(* IEC 61131-3 sources: daoli-st-library/DL_MathData (part 23) *)

(* ---- FC_DL_SearchMinMaxUdint.st ---- *)
(*
  ==================================================================
  组件名 Component  : FC_DL_SearchMinMaxUdint
  分类   Category   : DL_MathData
  复杂度 Complexity  : 低
  版本   Version    : 1.0.0
  功能   Purpose    : UDINT 域数组单遍扫描求最小值/最大值与双索引同出。前 nCount
                      个元素有效，一次循环同时出 uMin/uMax 与 uMinIdx/uMaxIdx
                      （首命中口径），无效哨兵按开关跳过并计数。
  来源   Source     : t2-1-lgf-math（LGF Math 极值检索族 UDINT 变体）
  溯源   Origin     : 极值检索属公开数学语义，clean-room 自研实现，未复制 LGF
                      或任何厂商私有库源码。
  平台   Platform   : 纯 IEC 61131-3（仅 FOR / 比较 / DINT_TO_UDINT），
                      CODESYS / TwinCAT / InoProShop / Machine Expert 通用
  分工声明 Split     : 与 FC_DL_SearchMinMax（LREAL 属主）及
                      FC_DL_SearchMinMaxDint（DINT 域同批连号件）三角互引——
                      本件为无符号域同构件，判式一律全序（<= / >=），不使用
                      任何减法比较（无符号域差值会回绕成大正数）。
  作者   Author     : 道莅代码库 · PLC 编程专家（R60）
  ------------------------------------------------------------------
  边界 Boundary     :
                      一 扫描个数钳位 1..4096，钳位置信息级码；
                      二 无效样本域：UDINT 域无 NaN，本件无效量定义为哨兵
                         DL_SMU_INVALID（= UDINT 最大位型 16#FFFF_FFFF），仅当
                         bIgnoreInvalid 为真时跳过（与 DINT 件哨兵取最小位型的
                         对称口径，头注释留痕）；
                      三 全量无效时 bValid = FALSE 且双索引回 0，不冒充 0 号位极值；
                      四 无符号比较只允许全序判式 <= / >=，禁用 a - b 差值判序；
                      五 无状态纯函数：每次调用局部量一律段 1 显式预置（R254）。
  接口偏离声明       : 派单示意 fMin/fMax（浮点命名），UDINT 输出按 R265 命名-类型
                      一致性落为 uMin/uMax，语义与引脚数一字不减。
  错误码   Codes    :
    16#0001_0604【信息级】计数越界已钳位（<1 早退，>4096 钳位续扫）
    16#0001_0605【信息级】无效哨兵样本已跳过，个数见 nSkipCnt
    16#0001_0606【故障级】全量无效，无有效极值，bValid = FALSE
  验收   Acceptance :
    算法已证（脚本）：未跑 ｜ 编译器已证（三平台）：未跑
    V1 数据 5 / 3 / 9 / 3，个数 4 → uMin=3 于索引 1，uMax=9 于索引 2
    V2 数据 16#FFFF_FFFE / 0 → uMin=0 于索引 1，uMax=16#FFFF_FFFE 于索引 0
    V3 哨兵 16#FFFF_FFFF 夹在有效值间，bIgnoreInvalid 真 → 跳过 1 个，码含 0605
    V4 个数 0 → bValid=FALSE、码 0604、双索引 0
    V5 全为哨兵且 bIgnoreInvalid 真 → bValid=FALSE、码 0606
  修订记录 Revision  :
    2026-11-21  v1.0.0  R60 首版（批 1 · 序号 2）
  ==================================================================
*)
FUNCTION FC_DL_SearchMinMaxUdint : BOOL
VAR_IN_OUT
    auValues : ARRAY[0..4095] OF UDINT; // 待扫描数组 [计数值]，前 nCount 个有效 / the scanned array, the first nCount entries valid
END_VAR
VAR_INPUT
    nCount         : DINT; // 有效样本数 [个]，钳位 1..4096 / the valid sample count, clamped to one through four thousand ninety six
    bIgnoreInvalid : BOOL; // 是否跳过无效哨兵值 [-] / whether the invalid sentinel entries are skipped
END_VAR
VAR_OUTPUT
    uMin     : UDINT; // 最小值 [计数值]，无有效样本时为 0 / the minimum value, zero when no valid sample
    uMax     : UDINT; // 最大值 [计数值]，无有效样本时为 0 / the maximum value, zero when no valid sample
    uMinIdx  : UDINT; // 最小值所在下标 [下标]，无有效样本时为 0 / the minimum index, zero when no valid sample
    uMaxIdx  : UDINT; // 最大值所在下标 [下标]，无有效样本时为 0 / the maximum index, zero when no valid sample
    nSkipCnt : UDINT; // 被跳过的无效哨兵个数 [个] / the skipped invalid sentinel count
    bValid   : BOOL;  // 结果是否有效（全量无效时为假）[-] / the result validity flag
    eErr     : UDINT; // 错误码，0 = 正常 / the error code, zero is ok
    bError   : BOOL;  // 错误标志，eErr 非 0 时为真 / the error flag, true when eErr is nonzero
END_VAR
VAR
    nI     : DINT;  // 扫描索引 [下标] / the scan index
    nUse   : DINT;  // 钳位后的扫描个数 [个] / the clamped scan count
    nSeen  : DINT;  // 已见有效样本数 [个] / the seen valid sample count
    uV     : UDINT; // 当前样本工作副本 [计数值] / the current sample working copy
    bHave  : BOOL;  // 已取得首个有效样本 [-] / the first valid sample taken flag
    bClamp : BOOL;  // 钳位发生标记 [-] / the clamp happened flag
END_VAR
VAR CONSTANT
    DL_SMU_DMAX    : DINT := 4096;          // 扫描个数上界 [个]，与数组容量一致 / the scan count bound aligned with the array capacity
    DL_SMU_INVALID : UDINT := 16#FFFF_FFFF; // 无效哨兵，等于 UDINT 最大位型（与 DINT 件取最小位型对称）/ the invalid sentinel equal to the UDINT maximum bit pattern
END_VAR

// 段 1｜返回值与错误状态预置安全值（四段式第一段，R45）+ 局部量显式预置（R254）/ segment 1, the preset of the return, the codes and the local guards
FC_DL_SearchMinMaxUdint := FALSE; // 返回值预置假 / preset the return false
uMin := 0; // 最小值预置零 / preset the minimum zero
uMax := 0; // 最大值预置零 / preset the maximum zero
uMinIdx := 0; // 最小索引预置零 / preset the minimum index zero
uMaxIdx := 0; // 最大索引预置零 / preset the maximum index zero
nSkipCnt := 0; // 跳过计数预置零 / preset the skipped count zero
bValid := FALSE; // 有效标志预置假（无有效样本前不宣称有效）/ preset the validity false
eErr := 16#0000_0000; // 错误码预置正常 / preset the code to ok
bError := FALSE; // 错误标志预置假 / preset the error flag false
nUse := 0; // 扫描个数预置零 / preset the scan count zero
nSeen := 0; // 有效样本数预置零 / preset the seen count zero
uV := 0; // 样本工作副本预置零 / preset the sample copy zero
bHave := FALSE; // 首样本标志预置假 / preset the first sample flag false
bClamp := FALSE; // 钳位标记预置假 / preset the clamp flag false

// 段 2｜扫描个数域闸（下界早退 + 上界钳位，边界一）/ segment 2, the scan count domain gate
IF nCount < 1 THEN // 低于下界，无样本可扫 / below the floor, nothing to scan
    eErr := 16#0001_0604; // 信息级：计数越界已钳位 / informational, the count clamped
    bError := TRUE; // 置错误标志（信息级随事件置位惯例）/ raise the error flag
    RETURN; // 早退：bValid 保持 FALSE，双索引保持 0 / early return with the validity false
END_IF
nUse := nCount; // 域内接管 / take the count inside the domain
IF nUse > DL_SMU_DMAX THEN // 高于上界 / above the bound
    nUse := DL_SMU_DMAX; // 钳到数组容量 / clamp to the array capacity
    bClamp := TRUE; // 置钳位标记 / raise the clamp flag
END_IF
IF bClamp THEN // 钳位发生时置信息级 / raise the informational code on a clamp
    eErr := 16#0001_0604; // 信息级：计数越界已钳位 / informational, the count clamped
    bError := TRUE; // 置错误标志 / raise the error flag
END_IF

// 段 3｜单遍扫描：首命中取极小与极大，索引与值同源写出（边界四）/ segment 3, the single pass scan with the first hit rule
FOR nI := 0 TO nUse - 1 DO // 有界循环（nUse 已钳 ≤4096）/ the bounded loop
    uV := auValues[nI]; // 取样本（索引已证在数组界内）/ take the sample, the index proven inside the bounds
    IF bIgnoreInvalid AND (uV >= DL_SMU_INVALID) THEN // 无效哨兵且开关为真（全序判式，不用等号）/ an invalid sentinel with the switch true, a total order test
        nSkipCnt := nSkipCnt + 1; // 跳过计数推进 / advance the skipped count
    ELSE // 有效样本参与极值 / a valid sample participates
        nSeen := nSeen + 1; // 有效样本数推进 / advance the seen count
        IF NOT bHave THEN // 首个有效样本：双向装填 / the first valid sample seeds both sides
            uMin := uV; // 最小值装填 / seed the minimum
            uMax := uV; // 最大值装填 / seed the maximum
            uMinIdx := DINT_TO_UDINT(nI); // 最小索引装填 / seed the minimum index
            uMaxIdx := DINT_TO_UDINT(nI); // 最大索引装填 / seed the maximum index
            bHave := TRUE; // 置首样本标志 / raise the first sample flag
        ELSE // 后续样本比较（首命中用严格判式，不覆盖等值）/ the later samples, strict tests keep the first hit
            IF uV < uMin THEN // 新极小 / a new minimum
                uMin := uV; // 更新最小值 / update the minimum
                uMinIdx := DINT_TO_UDINT(nI); // 更新最小索引（与值同源）/ update the minimum index from the same source
            ELSIF uV > uMax THEN // 新极大（uV ≥ uMin 前提下判极大即可，全序自证）/ a new maximum, proven by the total order
                uMax := uV; // 更新最大值 / update the maximum
                uMaxIdx := DINT_TO_UDINT(nI); // 更新最大索引（与值同源）/ update the maximum index from the same source
            END_IF
        END_IF
    END_IF
END_FOR

// 段 4｜结果复检兜底：全量无效判故障，信息级与故障级不共码（R258 三件套）/ segment 4, the result recheck
IF (nSeen > 0) AND (nSkipCnt > 0) AND (eErr = 16#0000_0000) THEN // 部分跳过且无先发事件 / a partial skip with no earlier event
    eErr := 16#0001_0605; // 信息级：无效哨兵样本已跳过 / informational, the invalid sentinels skipped
    bError := TRUE; // 置错误标志 / raise the error flag
END_IF
IF nSeen < 1 THEN // 无有效样本 / no valid sample
    eErr := 16#0001_0606; // 故障级：全量无效，无有效极值 / fault grade, no valid extremum
    bError := TRUE; // 置错误标志（R45 配对）/ raise the error flag, paired with the fault code
    bValid := FALSE; // 结果不可用 / the result void
    uMin := 0; // 双极值回安全值 / both extrema back to the safe zero
    uMax := 0; // 双极值回安全值 / both extrema back to the safe zero
    uMinIdx := 0; // 索引回 0（不冒充 0 号位极值，边界三）/ the index back to zero, not posing as the entry zero
    uMaxIdx := 0; // 索引回 0（不冒充 0 号位极值，边界三）/ the index back to zero, not posing as the entry zero
ELSE // 有有效样本 / with valid samples
    bValid := TRUE; // 结果有效 / the result is valid
    FC_DL_SearchMinMaxUdint := TRUE; // 返回成功 / return success
END_IF
END_FUNCTION

(* ---- FC_DL_SelEx.st ---- *)
(*
    FC_DL_SelEx —— 双通道选择泛型防御包装（REAL 域）
    ------------------------------------------------------------------
    分类      : DL_MathData / Sel
    前缀      : FC_DL_
    版本      : 1.0.0
    溯源      : IEC 61131-3 标准语义的道莅防御性实现
                （内部委托平台内建函数，外围统一错误码/钳位/双语文档；
                  未复制任何闭源厂商源码，参考实现仅限 MIT/Apache 许可）
    平台      : 纯 IEC 61131-3，CODESYS / TwinCAT / InoProShop 通用
    作者      : 道莅代码库 · PLC编程专家（R16）
    ------------------------------------------------------------------
    功能说明  : 双通道选择：bG=FALSE 选 fI0、bG=TRUE 选 fI1，选择运算用比较与
                IF/ELSE 实现（IEC SEL 语义），不重实现任何数学内核；
                选中通道非有限（NaN 或 ±INF）判为故障级 16#0001_02AC，返回 0.0 且 bValid=FALSE；
                未选中通道（备用通道）非有限仅置信息级 16#0001_01D4 记录，
                不影响本拍输出（输出仍为选中通道的有效值，bError=FALSE、bValid=TRUE）；
                选中与未选中同时异常时，故障级优先（返回 0.0）；
                ±INF 采用平台安全幅值比较判定（阈值高于 REAL 最大有限值 3.402823E38），NaN 用自不等判定；
                钳位方向：无钳位（故障拦截 / 信息记录，输出为通道原值或 0.0）。
    错误码    : 16#0001_02AC 选中通道非有限（NaN 或 ±INF）——故障级，返回 0.0
                16#0001_01D4 未选中通道（备用通道）非有限，仅记录——信息级，不影响本拍输出
                16#0001_01D5 预留禁用（信息级，不得挪用）
                16#0001_02AD 预留禁用（故障级，不得挪用）
                16#0001_02AE 预留禁用（故障级，不得挪用）
    状态机    : R6 标注 N/A —— 本组件为纯函数无顺序状态机，无 CASE 可写，非法状态不可能出现，故以本节说明替代 ELSE 兜底
    修订记录  : 2026-11-16 v1.0.0 首次入库（R16）
*)
FUNCTION FC_DL_SelEx : REAL
VAR_INPUT
    bG  : BOOL; // 选择输入，FALSE 选 fI0、TRUE 选 fI1 / select input, FALSE picks fI0, TRUE picks fI1
    fI0 : REAL; // 通道 0 输入 [无量纲] / channel 0 input
    fI1 : REAL; // 通道 1 输入 [无量纲] / channel 1 input
END_VAR
VAR_OUTPUT
    eErr   : UDINT; // 错误码，0=正常 / error id, 0=ok
    bError : BOOL;  // 是否出错，eErr 非 0 时为 TRUE / error flag, TRUE when eErr is nonzero
    bValid : BOOL;  // 输出是否有效可用 / output valid flag
END_VAR
VAR CONSTANT
    DL_REAL_INF_GUARD : LREAL := 4.0E38; // REAL 域 ±INF 判定阈值，高于 REAL 最大有限值 3.402823E38 [无量纲] / REAL +/-INF guard above max finite REAL 3.402823E38
END_VAR
VAR
    fSel      : REAL; // 选中通道值 [无量纲] / selected channel value
    bSelBad   : BOOL; // 选中通道非有限判定结果 / non-finite detection result of selected channel
    bIdleBad  : BOOL; // 未选中通道非有限判定结果 / non-finite detection result of unselected channel
END_VAR

// 段 1｜返回值与错误状态预置 / segment 1, preset return value and error status
FC_DL_SelEx := 0.0; // 故障缺省返回 0 [无量纲] / fault default returns 0
eErr   := 0;     // 预置无错误 / preset no error
bError := FALSE; // 预置无故障 / preset no fault
bValid := FALSE; // 预置无效，通过防御闸后置位 / preset invalid, set TRUE after guard passes

// 段 2｜通道选择与选中/未选中通道有限性判定 / segment 2, channel selection and finiteness check of both channels
IF bG THEN
    fSel := fI1; // TRUE 选通道 1 / TRUE picks channel 1
    bIdleBad := (fI0 <> fI0) OR (fI0 > DL_REAL_INF_GUARD) OR (fI0 < -DL_REAL_INF_GUARD); // 未选中通道 fI0 非有限判定 [无量纲] / unselected fI0 non-finite check
ELSE
    fSel := fI0; // FALSE 选通道 0 / FALSE picks channel 0
    bIdleBad := (fI1 <> fI1) OR (fI1 > DL_REAL_INF_GUARD) OR (fI1 < -DL_REAL_INF_GUARD); // 未选中通道 fI1 非有限判定 [无量纲] / unselected fI1 non-finite check
END_IF
bSelBad := (fSel <> fSel) OR (fSel > DL_REAL_INF_GUARD) OR (fSel < -DL_REAL_INF_GUARD); // 选中通道非有限判定（NaN 自不等 + 安全幅值判 ±INF） / selected channel non-finite check (NaN by self-inequality, +/-INF by safe magnitude)

// 段 3｜防御闸与输出（末段，故障级优先） / segment 3, guard and output (final, fault level first)
IF bSelBad THEN
    FC_DL_SelEx := 0.0;       // 故障级返回 0 [无量纲] / fault level returns 0
    eErr   := 16#0001_02AC;   // 选中通道非有限故障码 / selected channel non-finite fault id
    bError := TRUE;           // 置故障标志 / set fault flag
    bValid := FALSE;          // 输出无效 / output invalid
    RETURN;                   // 立即返回 / immediate return
ELSIF bIdleBad THEN
    FC_DL_SelEx := fSel;      // 输出选中通道原值，备用通道异常不影响本拍输出 / output selected value, idle channel anomaly does not affect this cycle
    eErr := 16#0001_01D4;     // 信息级：备用通道异常仅记录 / info level: idle channel anomaly recorded only
ELSE
    FC_DL_SelEx := fSel;      // 双通道均有限，正常输出选中值 / both channels finite, normal selected output
    eErr := 0; // 无错误 / no error
END_IF
bError := FALSE; // 信息级记录不置故障，故障分支已提前返回 / info-level record never raises fault, fault branch has returned
bValid := TRUE;  // 选中通道输出有效可用 / selected channel output is valid
END_FUNCTION

(* ---- FC_DL_SignedToUdintSat.st ---- *)
(*
  ==================================================================
  组件名 Component  : FC_DL_SignedToUdintSat
  分类   Category   : DL_MathData
  前缀   Naming     : FC_DL_ ｜ b/n/u/f/t/e/st 类型前缀制（R265）
  码位   Code ID    : 16#0001_0651（信息级）
  版本   Version    : 1.0.0
  复杂度 Complexity  : 低
  功能   Purpose    : DINT → UDINT 确定性转换：负值钳 0 并发信息级提示（多数平台此类
                      隐式转换行为不一，负值可能回绕成巨大正数，是 Modbus 寄存器打包的
                      经典故障源）。
  开源溯源 Origin    : IEC 61131-3 标准语义的道莅防御性实现（clean-room，无第三方代码行）
  许可证 License    : MIT
  参考   Reference  : IEC 61131-3:2013 §6.6.5 类型转换函数与 §6.5 有符号/无符号整数域定义
  平台   Platform   : 纯 IEC 61131-3（DINT_TO_UDINT / 比较），三平台通用
  依赖   Depends    : 仅 Standard.library（DINT_TO_UDINT 属标准转换函数）
  分工声明 Split     : FC_DL_UdintToDintChk 为反方向（UDINT → DINT，超上界钳 MAX 并置
                      故障级码），本件为 DINT → UDINT（负值钳零并置信息级码），两件成对，
                      边界互引（R216）。16 位入口（INT → UINT 同语义）按「禁新增同义邻件」
                      纪律并入本件重载，不另立文件。
  归属 Ownership     : 本件无 TYPE 声明，全部引脚为 IEC 标准原生类型。
  ------------------------------------------------------------------
  边界 Boundary     :
                      一 负值钳零是确定性合法行为而非故障：置信息级码、bValid 保持 TRUE、
                         bError 保持 FALSE（若按故障处理，Modbus 打包遇到合法的负温度
                         就会停机，分级明显错位）；
                      二 正域精确无溢出，域包含证明：DINT 非负域 [0, 2^31 − 1] 是全序
                         子集于 UDINT 全域 [0, 2^32 − 1]，即 [0, 2147483647] ⊂ [0, 4294967295]，
                         故 diIn ≥ 0 时 DINT_TO_UDINT 恒为精确映射，无须溢出分支；
                      三 反方向（UDINT → DINT）的越上界场景在本件域内不可能出现：
                         入参已是 UDINT 域内的值经 DINT 往返，属反方向件职责，本件不设分支；
                      四 纯函数：无记忆量、无定时器、无边沿实例，每调用重算。
  错误码 Codes      :
    16#0001_0651【信息级】负值已钳零（不锁存、不置 bError、bValid 保持 TRUE）
  验收 Acceptance   :
    算法已证（脚本）：未跑 ｜ 编译器已证（三平台）：未跑
    V1 0 → 0、bNegClamped = FALSE、无码
    V2 -1 → 0 + bNegClamped + 码 0651（bError = FALSE）
    V3 MIN（-2147483648）→ 0 + bNegClamped + 码 0651
    V4 MAX（2147483647）→ 2147483647 精确、无码
    V5 反方向向量（2^32−1 入 DINT）域上不可能，注释已给域包含关系，无须代码分支
  修订记录 Revision  :
    2026-11-21  v1.0.0  R62 首版（批 2 · 序号 6）
  ==================================================================
*)
FUNCTION FC_DL_SignedToUdintSat : BOOL
VAR_INPUT
    diIn : DINT; // 有符号输入 [−]，完整 DINT 域 / the signed input over the full DINT domain
END_VAR
VAR_OUTPUT
    udiOut      : UDINT; // 无符号结果 [−] / the unsigned result
    bNegClamped : BOOL;  // 负值已钳零 [-] / a negative value was clamped to zero
    bValid      : BOOL;  // 结果可用（本件恒 TRUE，保留引脚供族内统一）[-] / the result is usable, always true here
    eErr        : UDINT; // 错误码，0 = 正常 / the error code, zero is ok
    bError      : BOOL;  // 故障标志（本件只有信息级码，恒 FALSE）/ the fault flag, always false here since only an informational code exists
END_VAR
VAR CONSTANT
    DL_S2U_ZERO : DINT := 0;                  // 有符号零常量 [−] / the signed zero constant
    DL_S2U_UMIN : UDINT := 0;                 // 无符号零常量 [−] / the unsigned zero constant
    DL_S2U_DMAX : DINT := 2147483647;         // DINT 可表达上界 [−]，即 2^31−1 / the expressible DINT ceiling, two to the thirty first minus one
    DL_S2U_UMAX : UDINT := 4294967295;        // UDINT 可表达上界 [−]，即 2^32−1 / the expressible UDINT ceiling, two to the thirty second minus one
END_VAR

// 段 1｜返回值与全部出口预置安全值（R45 四段式第一段）/ segment 1, preset every outlet to its safe value
FC_DL_SignedToUdintSat := FALSE; // 返回值预置假 / preset the return false
udiOut := DL_S2U_UMIN; // 结果预置零 [−] / preset the result zero
bNegClamped := FALSE; // 负值钳零标志预置假 / preset the negative clamp flag false
bValid := FALSE; // 可用标志预置假，过闸后置位 / preset the validity false, raised after the gates
eErr := 16#0000_0000; // 错误码预置正常 / preset the code to ok
bError := FALSE; // 故障标志预置假（本件无故障级码）/ preset the fault flag false, no fault level code exists here

// 段 2｜负值钳零（边界一：确定性行为，非故障）/ segment 2, the negative clamp is a deterministic behaviour, not a fault
IF diIn < DL_S2U_ZERO THEN // 负值域 / the negative domain
    udiOut := DL_S2U_UMIN; // 钳零 [−] / clamp to zero
    bNegClamped := TRUE; // 置钳零标志 / raise the negative clamp flag
    eErr := 16#0001_0651; // 信息级：负值已钳零 / informational, a negative value was clamped to zero
    bError := FALSE; // 明确不置故障标志（信息级，R285 分级纪律）/ keep the fault flag false, this is informational
ELSE // 非负域：精确映射（边界二域包含证明）/ the non negative domain maps exactly
    udiOut := DINT_TO_UDINT(diIn); // 标准显式转换（DINT 非负域 ⊆ UDINT 全域）[−] / the standard explicit conversion, the signed non negative domain is a subset of the unsigned domain
END_IF

// 段 3｜统一出口（信息级钳零仍可用）/ segment 3, the unified outlet where a clamped zero stays usable
bValid := TRUE; // 负值钳零与正域精确均可用 / both the clamped zero and the exact positive domain are usable
FC_DL_SignedToUdintSat := TRUE; // 返回成功 / return success
END_FUNCTION

(* ---- FC_DL_SignumCalc.st ---- *)
(*
    FC_DL_SignumCalc —— 三态符号函数（浮点容差判零 + 非有限拦截）
    ------------------------------------------------------------------
    分类      : DL_MathData / Math-Sign
    前缀      : FC_DL_
    版本      : 1.0.0
    来源标签  : iec-std-wrapper（T0）
    溯源      : IEC 61131-3 标准语义的道莅防御性实现
                （纯比较逻辑，无内建数学内核依赖；未复制任何闭源厂商源码）
    平台      : 纯 IEC 61131-3，CODESYS / TwinCAT / InoProShop 通用
    分工声明  : 与存量 FC_DL_RealEqTolEx（判等）分工——EqTolEx 只回答是否相等，
                本件返回三态符号（负/零/正）；与 Hysteresis 分工——迟滞件带
                状态记忆，本件为无状态纯函数。
    作者      : 道莅代码库 · PLC 编程专家（R57）
    ------------------------------------------------------------------
    功能说明  : 返回输入的三态符号：|x| < fEps 判零返回 0（禁 = 判等）；
                x <= -fEps 返回 -1；x >= fEps 返回 +1。fEps <= 0 组态错误
                返回 0；非有限（NaN/Inf 双判据）返回 0 并出错误码。
    错误码    : 0000 正常 / 16#0003_0001 入参非有限 / 16#0003_0002 fEps 组态非法
    修订记录  : 2026-11-21 v1.0.0 首次入库（R57 批 3 · 序号 11）
*)
FUNCTION FC_DL_SignumCalc : INT
VAR_INPUT
    lrIn : LREAL;       // 输入实数 [工程单位] / input real value [engineering unit]
    fEps : LREAL := 1E-9; // 判零容差 [工程单位]，域 大于零 / the zero tolerance [engineering unit], above zero
END_VAR
VAR_OUTPUT
    eErr   : UDINT; // 错误码，0 = 正常 / error code, zero is ok
    bError : BOOL;  // 出错标志，eErr 非 0 时为真 / error flag, true when eErr is nonzero
    bValid : BOOL;  // 结果是否可用，拦截/组态错误时为假 / the result usable, false when intercepted
END_VAR

// 段 1｜返回值与错误状态预置安全值（四段式第一段，R45）/ segment 1, preset the return and error states
FC_DL_SignumCalc := 0; // 符号预置零 / preset the sign to zero
eErr   := 16#0000_0000; // 错误码预置正常 / preset the code to ok
bError := FALSE; // 错误标志预置假 / preset the error flag false
bValid := TRUE; // 有效标志预置真 / preset the valid flag true

// 段 2｜非有限拦截（双判据）：命中早退不比较 / segment 2, the non finite interception
IF (lrIn <> lrIn) OR ((lrIn - lrIn) <> (lrIn - lrIn)) THEN // NaN 或无穷 / NaN or infinity
    eErr   := 16#0003_0001; // 信息级：输入非有限返回零 / informational, a non finite input returns zero
    bError := TRUE; // 置错误标志 / raise the error flag
    bValid := FALSE; // 输出不可用 / the output void
    RETURN; // 返回预置安全值 0 / return the preset safe zero
END_IF

// 段 3｜组态闸：fEps <= 0 判组态错误（边界十一）/ segment 3, the config gate, a nonpositive tolerance illegal
IF (fEps <= 0.0) OR (fEps <> fEps) OR ((fEps - fEps) <> (fEps - fEps)) THEN // 容差非法或非有限 / an illegal or non finite tolerance
    eErr   := 16#0003_0002; // 错误级：容差组态非法 / error grade, an illegal tolerance config
    bError := TRUE; // 置错误标志 / raise the error flag
    bValid := FALSE; // 输出不可用 / the output void
    RETURN; // 返回预置安全值 0 / return the preset safe zero
END_IF

// 段 4｜三态符号判定：容差判零，禁 = 判等（边界十一）/ segment 4, the three state verdict with the tolerance
IF lrIn >= fEps THEN // 显著为正 / clearly positive
    FC_DL_SignumCalc := 1; // 返回正号 / return plus one
ELSIF lrIn <= -fEps THEN // 显著为负 / clearly negative
    FC_DL_SignumCalc := -1; // 返回负号 / return minus one
ELSE // 容差带内判零 / inside the tolerance band
    FC_DL_SignumCalc := 0; // 返回零 / return zero
END_IF
END_FUNCTION

(* ---- FC_DL_SimpsonQuad.st ---- *)
(*==============================================================================
 * 组件名称 (Component)  : FC_DL_SimpsonQuad
 * 所属子库 (Sublibrary) : DL_MathData
 * 当前版本 (Version)    : 1.0.0
 * 兼容性   (Platform)   : CODESYS 3.5+ / TwinCAT 3 / 汇川 InoProShop / 施耐德 Machine Expert
 *                         仅依赖 Standard.library（LOWER_BOUND / UPPER_BOUND / MOD），零厂商私有库
 * 功能描述 (Function)   : 复合辛普森 1/3 数值积分原语：对 n+1 个等距节点纵坐标（n 为偶数，
 *                         即节点数 >= 3 且区间数为偶）按公式
 *                           fI = fDx/3 × (aY[0] + 4×Σ奇节点 + 2×Σ偶内点 + aY[n])
 *                         单遍求积，返回积分值。适用功率-时间曲线求能、流量累计复核等
 *                         叶子级数值积分场景。
 * 接口     (Interface)  : 输入 aY 等距节点纵坐标数组（变长数组，按引传）、fDx 节点步长；
 *                         引用输出 bValid 有效标志（REFERENCE TO BOOL，当拍写回）；
 *                         返回值 = 积分值（bValid=FALSE 时返回 0）。
 * 边界     (Boundary)   : ① **属主边界（写死）：本件只做一次静态数组求积，不采样、不缓存、
 *                         不做时间触发**；采样与节点装载由调用方负责。
 *                         ② 奇偶判据用整数 MOD 2，禁浮点判奇偶。
 *                         ③ 拒算条件（任一成立返回 0 且 bValid=FALSE）：区间数 < 2（节点数
 *                         < 3）、区间数为奇数、fDx <= 容差、任一节点纵坐标非有限
 *                         （NaN 用自不等 x<>x 口径、Inf 用 (x-x)<>0 口径，R245）。
 *                         非有限值逐点前置剔除并**整体拒算**：部分积分结果不可信。
 *                         ④ 等距性由调用方保证（IN 语义声明）：本件不做步长一致性校验，
 *                         fDx 取相邻节点间距的名义值。
 *                         ⑤ 变长数组仅入 VAR_IN_OUT（IEC 61131-3 第 3 版对 ARRAY[*] 的
 *                         传参域限定），LOWER_BOUND/UPPER_BOUND 取实际上下界，不假设 0 起始。
 *                         ⑥ 零全局耦合（无 GVL / 无 VAR_EXTERNAL / 无物理地址）。
 * 分工声明 (Scope)      : 与 `FC_DL_PolyEvalHorner` 分工：多项式求值 ≠ 数值求积；与
 *                         `FC_DL_MultiPointLinear` 分工：分段线性插值 ≠ 积分。全库数值
 *                         积分原语由本件开族。
 * 来源标签 (Source Tag) : T2-1 LGF · Math 数学子族（公开数学定义 clean-room，复合辛普森
 *                         1/3 法则为教科书公开公式，零代码行复制）
 * 码表     (Codes)      : 本件不占用任何全局数字码位。出口为 LREAL 积分值 + BOOL 有效标志；
 *                         数字码位待主控收口阶段统一派号。
 * 红线自检 (Redline)    : R1 ✓ 零 GVL/VAR_EXTERNAL ｜ R2 ✓ 零 %I/%Q/%M ｜ R3 ✓ 纯 IEC 61131-3
 *                         R4 ✓ 步长容差闸 + 非有限前置剔除 + 奇偶整数判据 ｜ R5 ✓ 声明逐行同行双语注释
 *                         R6 N/A（纯函数无状态机） ｜ R7 N/A（无实例调用）
 * 修订历史 (Revision)   : 2026-11-20  v1.0.0  R48 首版（批次 1 · 序号 2）
 *                         验收向量：3 节点 y=[0,1,0]、dx=1 → 4/3；4 节点（奇区间数）拒算；
 *                         含 NaN 节点整体拒算；dx=0 拒算。
 *==============================================================================*)

FUNCTION FC_DL_SimpsonQuad : LREAL
VAR_IN_OUT
    aY : ARRAY[*] OF LREAL;    // 等距节点纵坐标数组（长度 n+1，n 偶），单位随被积量 [被积量纲] / Ordinates at equidistant nodes
END_VAR
VAR_INPUT
    fDx    : LREAL;                 // 节点步长，域 > 容差；等距性由调用方保证（IN 语义） [横轴单位] / Node spacing, > epsilon, uniformity by caller
    bValid : REFERENCE TO BOOL;     // 有效标志（引用传参；FALSE=拒算） [-] / Validity flag, by-reference, FALSE when rejected
END_VAR
VAR
    nLo  : DINT;                    // 数组实际下界索引 / Actual lower array index
    nHi  : DINT;                    // 数组实际上界索引 / Actual upper array index
    nInt : DINT;                    // 区间数 = 节点数 - 1，须为正偶数 / Interval count, positive even
    i    : DINT;                    // 求和循环索引 / Summation loop index
    fSum : LREAL;                   // 括号内加权和中间量 / Weighted sum accumulator
END_VAR
VAR CONSTANT
    DL_SQ_EPS : LREAL := 1.0E-12;   // 步长判零容差 [横轴单位] / Spacing zero epsilon
    DL_SQ_W4  : LREAL := 4.0;       // 辛普森奇节点权重 [-] / Simpson odd-node weight
    DL_SQ_W2  : LREAL := 2.0;       // 辛普森偶内点权重 [-] / Simpson even-interior weight
    DL_SQ_W3  : LREAL := 3.0;       // 1/3 法则除数 [-] / Divisor of the one-third rule
END_VAR

bValid := FALSE;                                       // 缺省拒算 / Default: invalid
FC_DL_SimpsonQuad := 0.0;                              // 拒算返回 0 / Rejected returns zero
nLo  := LOWER_BOUND(aY, 1);                            // 取实际下界，不假设 0 起始 / Actual lower bound, no zero assumption
nHi  := UPPER_BOUND(aY, 1);                            // 取实际上界 / Actual upper bound
nInt := nHi - nLo;                                     // 区间数 / Interval count
IF (nInt < 2) OR ((nInt MOD 2) <> 0) OR (fDx <= DL_SQ_EPS) THEN
    RETURN;                                            // 区间数不足 / 奇区间数 / 步长非正：拒算（整数奇偶判据）/ Too few or odd intervals or bad spacing: reject
END_IF
FOR i := nLo TO nHi DO
    IF (aY[i] <> aY[i]) OR ((aY[i] - aY[i]) <> 0.0) THEN
        RETURN;                                        // 任一节点非有限（NaN 自不等 / Inf 差非零）：整体拒算（R245）/ Any non-finite node: reject wholly
    END_IF
END_FOR

fSum := aY[nLo] + aY[nHi];                             // 两端节点权重 1 / End nodes carry weight one
FOR i := (nLo + 1) TO (nHi - 1) DO
    IF ((i - nLo) MOD 2) <> 0 THEN
        fSum := fSum + DL_SQ_W4 * aY[i];               // 奇节点权重 4 / Odd nodes weight four
    ELSE
        fSum := fSum + DL_SQ_W2 * aY[i];               // 偶内点权重 2 / Even interior nodes weight two
    END_IF
END_FOR

FC_DL_SimpsonQuad := fSum * fDx / DL_SQ_W3;            // 除数为常量 3，无除零 / Constant divisor three, no zero division
bValid := TRUE;                                        // 求积有效 / Result valid

END_FUNCTION

(* ---- FC_DL_SincSafe.st ---- *)
(*==============================================================================
 * 名称 : FC_DL_SincSafe —— 安全 sinc(x)=sin(x)/x（0 点泰勒展开防除零）
 * 分类 / 前缀 / 版本 : DL_MathData / FC_DL_ / 1.0.0
 * 溯源 : 开源语义参考（OSCAT/AixOCAT 族，MIT）或 clean-room IEC 实现，未复制源码
 * 平台 : 纯 IEC 61131-3
 * 功能说明 : 计算 sinc(x)=sin(x)/x。|x|<1.0E-8 时用四阶泰勒近似
 *            1 - x^2/6 + x^4/120（该区间误差 < 1.0E-16 量级），避免 0 点
 *            除零；其余区间直接 sin(x)/x（|x|>=1.0E-8 保证分母非零）。
 *            边界处理：输入非有限（NaN/±Inf）置 eErr 返回 0.0；x=0 精确落
 *            入泰勒支路返回 1.0（sinc 极限值），属正确结果非故障。
 * 错误码 : 16#0001_1B0F = 输入非有限（NaN/±Inf）
 *          eErr=0 且 bValid=TRUE 表示返回值可用
 * 状态机 : R6 标注 N/A（纯函数无顺序状态，以本节替代 ELSE 兜底）
 * 红线 : R1/R2/R3 ✓ 零全局/零IO/纯IEC ｜ R4 ✓ 非有限拦截/除零防护 ｜ R10 ✓ 标准转换 ｜ R11 ✓ 分号收尾 ｜ R15 ✓ 无保留字撞名
 * 修订记录 : 2026-11-23 v1.0.0 首次入库（R76）
 *============================================================================*)
FUNCTION FC_DL_SincSafe : LREAL
VAR_INPUT
    fX : LREAL;    // 输入自变量 [rad] / input argument in radians
END_VAR
VAR_OUTPUT
    eErr   : UDINT;    // 故障码，0=正常，1B0F=输入非有限 / error code
    bError : BOOL;     // TRUE=本件发生故障 / TRUE when fault occurred
    bValid : BOOL;     // TRUE=返回值可用 / TRUE when return value is usable
END_VAR
VAR
    _x2 : LREAL;       // x 的平方（泰勒中间量）/ squared input for Taylor series
    _x4 : LREAL;       // x 的四次方（泰勒中间量）/ fourth power for Taylor series
END_VAR

FC_DL_SincSafe := 0.0;                       // 返回值预设 0.0 / preset return to zero
eErr   := 16#0000_0000;                      // 故障码清零 / clear error code
bError := FALSE;                             // 故障标志清零 / clear error flag
bValid := TRUE;                              // 预设输出可用 / preset valid flag

IF (fX <> fX) OR ((fX - fX) <> (fX - fX)) THEN    // NaN 或 ±Inf / NaN or infinite
    eErr   := 16#0001_1B0F;                  // 置非有限故障码 / set non-finite code
    bError := TRUE;                          // 置故障标志 / set error flag
    bValid := FALSE;                         // 返回值不可用 / return not usable
    RETURN;                                  // 返回 0.0 / return zero
END_IF

IF ABS(fX) < 1.0E-8 THEN                     // 0 点邻域走泰勒支路 / Taylor branch near zero
    _x2 := fX * fX;                          // 平方中间量 / square
    _x4 := _x2 * _x2;                        // 四次方中间量 / fourth power
    FC_DL_SincSafe := 1.0 - _x2 / 6.0 + _x4 / 120.0;    // 四阶泰勒近似（0 点返回 1.0）/ 4th-order Taylor
ELSE                                         // 非零区间直接作商（分母 |x|>=1E-8 非零）/ direct quotient
    FC_DL_SincSafe := SIN(fX) / fX;          // sin(x)/x，分母已保证非零 / denominator guaranteed nonzero
END_IF

END_FUNCTION

(* ---- FC_DL_SinDeg.st ---- *)
(*==============================================================================
 * 名称 : FC_DL_SinDeg —— 角度制正弦（度入参，弧度内部换算）
 * 分类 / 前缀 / 版本 : DL_MathData / FC_DL_ / 1.0.0
 * 溯源 : 开源语义参考（OSCAT/AixOCAT 族，MIT）或 clean-room IEC 实现，未复制源码
 * 平台 : 纯 IEC 61131-3
 * 功能说明 : 返回 sin(fDeg)：内部换算弧度 fDeg * PI / 180 后调用标准 SIN，
 *            PI 取 LREAL 字面量 3.14159265358979323846（双精度最近舍入）。
 *            边界处理：输入非有限（NaN：f<>f；±Inf：(f-f)<>(f-f)）置 eErr
 *            返回 0.0；|fDeg|>1.0E12 时大角换算精度塌陷，同置 eErr 返回 0.0。
 * 错误码 : 16#0001_1B09 = 输入非有限（NaN/±Inf）或角度量超安全量程 ±1.0E12
 *          eErr=0 且 bValid=TRUE 表示返回值可用
 * 状态机 : R6 标注 N/A（纯函数无顺序状态，以本节替代 ELSE 兜底）
 * 红线 : R1/R2/R3 ✓ 零全局/零IO/纯IEC ｜ R4 ✓ 非有限拦截/量程防护 ｜ R10 ✓ 标准转换 ｜ R11 ✓ 分号收尾 ｜ R15 ✓ 无保留字撞名
 * 修订记录 : 2026-11-23 v1.0.0 首次入库（R76）
 *============================================================================*)
FUNCTION FC_DL_SinDeg : LREAL
VAR_INPUT
    fDeg : LREAL;    // 输入角 [度] / input angle in degrees
END_VAR
VAR_OUTPUT
    eErr   : UDINT;    // 故障码，0=正常，1B09=输入非有限或超量程 / error code
    bError : BOOL;     // TRUE=本件发生故障 / TRUE when fault occurred
    bValid : BOOL;     // TRUE=返回值可用 / TRUE when return value is usable
END_VAR

FC_DL_SinDeg := 0.0;                         // 返回值预设 0.0 / preset return to zero
eErr   := 16#0000_0000;                      // 故障码清零 / clear error code
bError := FALSE;                             // 故障标志清零 / clear error flag
bValid := TRUE;                              // 预设输出可用 / preset valid flag

IF (fDeg <> fDeg) OR ((fDeg - fDeg) <> (fDeg - fDeg))    // NaN 或 ±Inf / NaN or infinite
   OR (ABS(fDeg) > 1.0E12) THEN              // 超安全量程（精度塌陷防护）/ beyond safe range
    eErr   := 16#0001_1B09;                  // 置故障码 / set error code
    bError := TRUE;                          // 置故障标志 / set error flag
    bValid := FALSE;                         // 返回值不可用 / return not usable
    RETURN;                                  // 返回 0.0 / return zero
END_IF

FC_DL_SinDeg := SIN(fDeg * 3.14159265358979323846 / 180.0);    // 度转弧度后取正弦 / degrees to radians, then sine

END_FUNCTION

(* ---- FC_DL_SinEx.st ---- *)
(*
    FC_DL_SinEx —— 正弦防御包装（2π 周期归约保精度 + 非有限拦截 + 超大角度降级）
    ------------------------------------------------------------------
    分类      : DL_MathData / Math-Trig
    前缀      : FC_DL_
    版本      : 1.0.0
    溯源      : IEC 61131-3 标准语义的道莅防御性实现
                （内部委托平台内建函数，外围统一错误码/钳位/双语文档；
                  未复制任何闭源厂商源码，参考实现仅限 MIT/Apache 许可）
    平台      : 纯 IEC 61131-3，CODESYS / TwinCAT / InoProShop 通用
    作者      : 道莅代码库 · PLC编程专家（R15）
    ------------------------------------------------------------------
    功能说明  : 求输入弧度的正弦值。入口先做非有限拦截（NaN/Inf 返回 0.0
                并置 16#0001_0163）；随后按 2π 做周期归约，商取 FLOOR 语义避免负向
                误差，商绝对值 < 2.0E9 保证 DINT 转换不溢出；超大角度
                （绝对值 > 1.0E12 或商超 DINT 安全域）降级处理：置 16#0001_0163、
                bValid=FALSE 但仍继续计算；域内委托内建 SIN，结果再做
                NaN 复检兜底，全程不输出 NaN/Inf。
    错误码    : 0000 正常 / 16#0001_0163 入参越界（非有限输入或超大角度降级，已归零/降级可用）
    修订记录  : 2026-11-16 v1.0.0 首次入库（R15）
*)
FUNCTION FC_DL_SinEx : LREAL
VAR_INPUT
    lrRad : LREAL; // 输入角度 [rad]，任意有限弧度值 / input angle [rad], any finite radian value
END_VAR
VAR_OUTPUT
    eErr : UDINT; // 错误码，0=正常，1=入参越界（非有限或超大角度） / error id, 0=ok, 1=input out of domain (non-finite or super-large angle)
    bError   : BOOL; // 是否出错，eErr 非 0 时为 TRUE / error flag, TRUE when eErr is nonzero
    bValid   : BOOL; // 输出是否有效可用，超大角度降级时为 FALSE / output valid, FALSE for degraded super-large angle
END_VAR
VAR
    lrQ   : LREAL; // 周期商 [周期数]，输入角除以 2π / cycle quotient [cycles], input divided by two pi
    nCyc  : DINT; // 归约周期数 [周期数]，FLOOR 语义整数 / reduction cycle count [cycles], integer with floor semantics
    lrRed : LREAL; // 归约后弧度 [rad]，域约至 0 到 2π / reduced angle [rad], bounded to 0 to 2 pi
END_VAR
VAR CONSTANT
    DL_SN_MAXREAL : LREAL := 1.7976931348623157E308; // 双精度有限极值 [rad]，超界判无穷 / double precision finite max [rad], beyond treated as infinity
    DL_SN_TWOPI   : LREAL := 6.283185307179586; // 圆周率两倍 [rad]，归约模数 / two pi [rad], reduction modulus
    DL_SN_BIG     : LREAL := 1.0E12; // 超大角度阈值 [rad]，超过判降级 / super-large angle threshold [rad], beyond degraded
    DL_SN_QMAX    : LREAL := 2.0E9; // 周期商安全域 [周期数]，保证 DINT 转换不溢出 / quotient safe bound [cycles], keeps DINT conversion overflow-free
    DL_SN_EPS     : LREAL := 1.0E-9; // 浮点容差 [无量纲] / floating point tolerance [dimensionless]
END_VAR

// 段 1｜返回值与错误状态预置，任何早退路径不留脏码 / segment 1, preset return value and error states
FC_DL_SinEx := 0.0; // 返回值预置安全值 0.0 / preset return to safe value 0.0
eErr    := 16#0000_0000; // 错误码预置正常 / preset error id to ok
bError      := FALSE; // 错误标志预置无错 / preset error flag to FALSE
bValid      := TRUE; // 有效标志预置可用 / preset valid flag to TRUE

// 段 2｜非有限拦截：NaN 用自不等判据，无穷用超极值判据 / segment 2, non-finite interception
IF (lrRad <> lrRad) OR (lrRad > DL_SN_MAXREAL) OR (lrRad < -DL_SN_MAXREAL) THEN
    eErr := 16#0001_0163; // 信息级：输入非有限，已归零 / informational, non-finite input, zeroed
    bError   := TRUE; // 置错误标志 / raise error flag
    bValid   := FALSE; // 输出不可用 / output invalid
    RETURN; // 返回预置安全值 0.0 / return preset safe value 0.0
END_IF

// 段 3｜2π 周期归约（FLOOR 语义）：商超 DINT 安全域则跳过归约原值直通 / segment 3, two-pi reduction with floor semantics, skipped when quotient exceeds the DINT safe bound
lrQ := lrRad / DL_SN_TWOPI; // 周期商 [周期数] / cycle quotient [cycles]
IF ABS(lrQ) < DL_SN_QMAX THEN
    nCyc := TRUNC(lrQ); // 向零截取周期数 / truncate quotient toward zero
    IF (lrQ < 0.0) AND (ABS(lrQ - DINT_TO_LREAL(nCyc)) > DL_SN_EPS) THEN
        nCyc := nCyc - 1; // 负非整数商补一，落实 FLOOR 语义 / decrement for negative non-integer quotient to enforce floor semantics
    END_IF
    lrRed := lrRad - DL_SN_TWOPI * DINT_TO_LREAL(nCyc); // 归约后弧度 [rad] / reduced angle [rad]
ELSE
    lrRed := lrRad; // 商超安全域，放弃归约原值直通 / quotient beyond safe bound, reduction skipped
END_IF

// 段 4｜超大角度精度闸：置 16#0001_0163 降级但继续计算 / segment 4, super-large angle precision gate, degraded with code 1 but computation continues
IF (ABS(lrRad) > DL_SN_BIG) OR (ABS(lrQ) >= DL_SN_QMAX) THEN
    eErr := 16#0001_0163; // 信息级：超大角度，精度不可保证 / informational, super-large angle, precision not guaranteed
    bError   := TRUE; // 置错误标志 / raise error flag
    bValid   := FALSE; // 降级输出，需上层注意 / degraded output, upper layer attention required
END_IF

// 段 5｜委托内建 SIN + 结果 NaN 复检兜底 / segment 5, delegation to built-in SIN with result NaN recheck
FC_DL_SinEx := SIN(lrRed); // 委托内建 SIN 内核，不自实现三角内核 / delegate to built-in SIN kernel
IF FC_DL_SinEx <> FC_DL_SinEx THEN
    FC_DL_SinEx := 0.0; // 兜底安全值 / bottom-line safe value
    IF eErr = 16#0000_0000 THEN
        eErr := 16#0001_0163; // 首事件优先置码 / first-event priority code
        bError   := TRUE; // 置错误标志 / raise error flag
        bValid   := FALSE; // 输出不可用 / output invalid
    END_IF
END_IF
END_FUNCTION

(* ---- FC_DL_SinterShrinkageCalc.st ---- *)
(*
  Component : FC_DL_SinterShrinkageCalc
  Category  : DL_MathData
  Type      : FC
  Complexity: C1
  VERSION   : v1.0.0
  功能      : 烧结线收缩率与模具尺寸补偿：按烧结前后密度比开立方得线收缩率，并由成品尺寸反算所需模具尺寸。
  开源溯源  : 道莅原创 clean-room 自研（无外部代码引用）｜License: MIT
  边界条件  : ① 生坯密度与烧结密度均须 > 1e-9（均为除子），否则返回哨兵 -1；
              ② 烧结密度低于生坯密度时收缩率为负（膨胀），照实输出不钳位，便于诊断工艺异常；
              ③ 反算模具尺寸用 成品尺寸 / 线性比例因子，比例因子为 0 时不计算。
*)
FUNCTION FC_DL_SinterShrinkageCalc : REAL
VAR_INPUT
    fGreenDensGcm3 : REAL;   (* 烧结前生坯密度 [g/cm³] Green density before sintering *)
    fSinterDensGcm3: REAL;   (* 烧结后密度 [g/cm³] Sintered density *)
    fFinalDimMm    : REAL;   (* 成品目标尺寸 [mm] Final part dimension *)
END_VAR
VAR_OUTPUT
    fLinFactor  : REAL;   (* 线性比例因子（成品/模具） [-] Linear scale factor *)
    fShrinkPct  : REAL;   (* 线收缩率 [%] Linear shrinkage percent *)
    fDieDimMm   : REAL;   (* 反算模具尺寸 [mm] Die dimension *)
    xValid      : BOOL;   (* 计算有效性标志 [-] Calculation valid flag *)
END_VAR
VAR CONSTANT
    DL_EPS      : REAL := 1.0E-9;   (* 除零判定容差 [无量纲] Divide-by-zero tolerance *)
    DL_THIRD    : REAL := 0.3333333333333333;  (* 立方根指数 [-] Cube-root exponent *)
    DL_PCT_BASE : REAL := 100.0;    (* 百分比基准 [%] Percent base *)
    DL_ONE      : REAL := 1.0;      (* 单位常数 [-] Unity constant *)
END_VAR
(* 出口预置：三出口统一预置 *)
fLinFactor := 1.0; fShrinkPct := 0.0; fDieDimMm := 0.0; xValid := FALSE;
(* 非有限拦截：自反判 NaN，自身差值判 Inf *)
IF (fGreenDensGcm3 <> fGreenDensGcm3) OR ((fGreenDensGcm3 - fGreenDensGcm3) <> 0.0)
   OR (fSinterDensGcm3 <> fSinterDensGcm3) OR ((fSinterDensGcm3 - fSinterDensGcm3) <> 0.0)
   OR (fFinalDimMm <> fFinalDimMm) OR ((fFinalDimMm - fFinalDimMm) <> 0.0) THEN
    FC_DL_SinterShrinkageCalc := -1.0;  (* 哨兵 -1：输入非有限 / Sentinel -1 non-finite *)
    RETURN;
END_IF
(* 组态域闸：两个密度均为除子，成品尺寸须为正 *)
IF (fGreenDensGcm3 <= DL_EPS) OR (fSinterDensGcm3 <= DL_EPS) OR (fFinalDimMm <= DL_EPS) THEN
    FC_DL_SinterShrinkageCalc := -1.0;  (* 哨兵 -1：组态非法 / Sentinel -1 bad config *)
    RETURN;
END_IF
(* 质量守恒：体积比 = 密度比的反比，线比例因子 = 体比例因子的立方根 *)
fLinFactor := EXPT(fGreenDensGcm3 / fSinterDensGcm3, DL_THIRD);
(* 线收缩率：收缩为正，膨胀为负，照实输出便于工艺诊断 *)
fShrinkPct := (DL_ONE - fLinFactor) * DL_PCT_BASE;
(* 反算模具尺寸：成品 = 模具 × 线比例因子，因子为 0 时不下发 *)
IF fLinFactor > DL_EPS THEN
    fDieDimMm := fFinalDimMm / fLinFactor;
END_IF
xValid := TRUE;                            (* 链路有效 / Chain valid *)
FC_DL_SinterShrinkageCalc := fShrinkPct;   (* 返回线收缩率 [%] / Return linear shrinkage *)
END_FUNCTION

(* ---- FC_DL_SlewRateCalc.st ---- *)
(*
  ==================================================================
  组件名 Component  : FC_DL_SlewRateCalc
  分类   Category   : DL_MathData
  前缀   Naming     : FC_DL_ ｜ b/n/u/f 类型前缀制（R265）
  版本   Version    : 1.0.0
  功能   Purpose    : 采样间变化率：fRate = (fCurVal − fPrevVal) / fDtSec
                      [工程单位/s]。fDtSec ≤ 0 闸（除法前置，含容差判零
                      语义：≤0 即拒）；输入非有限闸；差值/结果非有限复
                      核（有限大数相减可溢出 Inf）。纯无状态函数，采样
                      时刻由调用方维护（前后两次采样值由调用方快照传入），
                      本件不驻留上拍数据。
  来源   Source     : t2-1-lgf-technology（差分变化率为公开数值口径，
                      实现零源码复制）
  互引   Cross-ref  : FB_DL_CycleTimeMeasure（同族周期测量件：其扫描周期
                      口径可作 fDtSec 注入来源）；FC_DL_NormTo01（同族
                      数学原子邻件）
  平台   Platform   : 纯 IEC 61131-3 四则 + ABS，三平台通用
  依赖   Depends    : 无 DL_ 内部依赖；无标准库
  红线   Redline    : R1 零全局/VAR_EXTERNAL/R2 零 %I/%Q/R3 纯 IEC 标准
                      R4 除零闸（dt ≤ 0 前置）+ 非有限三面闸（输入/差值/
                      结果）/R5 全变量双语同行注释/R6 纯函数无状态机
                      （CASE 不适用）/R7 无定时器与沿检测/R8 容差常量化
  错误码 Codes      : 01【失效级】采样间隔非法（fDtSec ≤ 0），返回 0
                      02【失效级】任一输入非有限（NaN 自反判 / Inf 上限
                      兜底判）或差值/结果非有限，返回 0
  码位反证 Note     : 01/02 分立依据（R90）：01 在时基面（调用方采样节拍
                      组态/断拍）、02 在数据面可观测；02 若并入 01，则
                      「时基正常仍失败」的数据病态将不可观测，故必须分立。
  验收   Acceptance : V1 10→12 / dt=0.5s → 4 [u/s] ｜ V2 dt=0 → 码 01
                      ｜ V3 dt=−1 → 码 01 ｜ V4 含 NaN → 码 02 ｜
                      V5 1E308→−1E308 / dt=1 → 码 02（差值 Inf）
  变更   Revision   : 2026-11-22  v1.0.0  R67 首版（编码阶段批 2 序 4）
  ==================================================================
*)
FUNCTION FC_DL_SlewRateCalc : LREAL
VAR_INPUT
    fCurVal  : LREAL;  // 当前采样值 [工程单位] / the current sample value
    fPrevVal : LREAL;  // 前一采样值（调用方快照）[工程单位] / the previous sample value, snapshot by the caller
    fDtSec   : LREAL;  // 采样间隔 [s]，须 > 0 / the sample interval in seconds, must be positive
END_VAR
VAR_OUTPUT
    bValid : BOOL;     // 变化率可用标志 [-] / the slew rate usable flag
    nErrId : UDINT;    // 错误码，0=正常，01/02 见头注 [码] / the error code [code]
END_VAR
VAR
    fDelta : LREAL;    // 差值工作寄存器 [工程单位] / the delta working register
END_VAR
VAR CONSTANT
    SRC_FIN_MAX  : LREAL := 1.7976931348623157E308; // LREAL 有限上限 / the finite LREAL limit
    SRC_ERR_NONE : UDINT := 16#0000_0000;           // 无错误 [码] / no error [code]
    SRC_ERR_DT   : UDINT := 16#0000_0001;           // 码 01：采样间隔非法 / code 01, illegal interval
    SRC_ERR_NAN  : UDINT := 16#0000_0002;           // 码 02：非有限 / code 02, non finite
END_VAR

// 段 1｜输出预置 / segment 1, preset the outputs
FC_DL_SlewRateCalc := 0.0;  // 失效缺省返回 0 / fault default returns zero
bValid := FALSE;            // 预置不可用 / preset unusable
nErrId := SRC_ERR_NONE;     // 预置无错误 / preset no error

// 段 2｜采样间隔闸（码 01）：除法前置，≤0 即拒（含 dt 非有限：NaN 与任何
//      比较为 FALSE，会漏闸，故先自反判）/ segment 2, the interval gate
IF (fDtSec <> fDtSec) OR (fDtSec <= 0.0) THEN
    nErrId := SRC_ERR_DT;   // 时基面失效 / the time base failure
    RETURN;
END_IF

// 段 3｜输入非有限闸（码 02）/ segment 3, the input finite gate
IF (fCurVal <> fCurVal) OR (fPrevVal <> fPrevVal)
   OR (ABS(fCurVal) > SRC_FIN_MAX) OR (ABS(fPrevVal) > SRC_FIN_MAX) OR (ABS(fDtSec) > SRC_FIN_MAX) THEN
    nErrId := SRC_ERR_NAN;
    RETURN;
END_IF

// 段 4｜差分与除法（分母 = fDtSec，段 2 已闸）/ segment 4, the delta and the division
fDelta := fCurVal - fPrevVal;             // 差值 [工程单位] / the delta
IF (fDelta <> fDelta) OR (ABS(fDelta) > SRC_FIN_MAX) THEN
    nErrId := SRC_ERR_NAN;                // 有限差溢出 Inf 兜底 / the delta overflow fallback
    RETURN;
END_IF
FC_DL_SlewRateCalc := fDelta / fDtSec;    // 变化率 [工程单位/s] / the slew rate
IF (FC_DL_SlewRateCalc <> FC_DL_SlewRateCalc) OR (ABS(FC_DL_SlewRateCalc) > SRC_FIN_MAX) THEN
    nErrId := SRC_ERR_NAN;                // 结果非有限复核 / the result finiteness recheck
    FC_DL_SlewRateCalc := 0.0;            // 失效回缺省 0 / fault default zero
    RETURN;
END_IF
bValid := TRUE;                           // 变化率可用 / the slew rate is usable
END_FUNCTION

(* ---- FC_DL_SolarPositionCalc.st ---- *)
(*==============================================================================
 * 组件名称 (Component)  : FC_DL_SolarPositionCalc
 * 所属子库 (Sublibrary) : DL_MathData
 * 当前版本 (Version)    : 1.0.0
 * 兼容性   (Platform)   : CODESYS 3.5 / TwinCAT 3 / 汇川 InoProShop / Machine Expert
 *                         仅依赖 Standard.library（SIN / COS / TAN / ASIN / ATAN2 / ABS / LIMIT）
 * 功能描述 (Function)   : 由本地标准时（年 / 月 / 日 / 时 / 分）、纬度、经度与时区偏移，
 *                         按 NOAA 公开的简化天文算法求太阳赤纬、均时差、真太阳时、时角、
 *                         高度角与方位角。现场用途：光伏跟踪支架逆跟踪角、建筑遮阳帘、
 *                         日光温室补光窗口、日照辐射计的姿态修正。
 *                         方位角约定：正北 0 度、顺时针递增（东 90、南 180、西 270）。
 *                         天顶约定：高度角高于 89.5 度（或高度角余弦小于 0.00873）时，
 *                         方位角在物理上不可辨，本件统一置 180.0 度（正南）并保持该约定不变，
 *                         上层如另有偏好须在调用侧追加判别，不得依赖本件给出「就近方位」。
 * 出口契约 (Exit)       : 函数返回值 = 太阳高度角（与出口 fElevation 同值）；输入域外一律
 *                         返回 0.0 且 bValid = FALSE，绝不输出「看起来合理」的错值。
 * 开源溯源 (Origin)     : 来源标签 lgf-datetimer。许可证：LGF 为免费闭源发布，未取得源码，
 *                         不构成衍生作品。借鉴点仅为「Date and Timer 组把日历天数、周数、
 *                         天文钟、多段定时并列」的分类骨架，以及天文钟「本地时间 + 经纬度
 *                         求太阳位置」的参数域划分。全部公式取 NOAA 公开算法（公共领域），
 *                         实现、常量、归一策略、域守护与错误码 100% clean-room 自有。
 * 码位说明 (Codes)      : 信息级 16#0001_0136（年月时分 / 经纬度 / 时区域外）/
 *                         16#0001_0137（日超出当月实际天数，含闰年判定）。共 2 码，
 *                         落在 R12 计划第 1.2 节本件码段内，无段外码。
 * 依赖     (Depends)    : 无 DL_ 内部依赖；Standard.library 三角函数与 LIMIT
 * 红线自检 (Redline)    : 1 ✓ 零全局变量表依赖、零外部变量声明、零物理地址
 *                         2 ✓ 纯 IEC 61131-3，无指针、无厂商库
 *                         3 ✓ 经纬度与时区域外早退、ASIN 入参钳位、ATAN2 双零守护、
 *                             时角与方位角归一用条件加减（不用 MOD）、循环带守卫
 *                         4 ✓ 全变量中英双语同行注释
 *                         5 N/A 纯函数无状态机 ｜ 6 N/A 无定时器与边沿实例
 *                         7 ✓ END_FUNCTION 位于文件最后有效行
 * 算法出处与精度声明    :
 *   NOAA Solar Calculator 公开的傅里叶级数（赤纬 7 项、均时差 5 项），
 *   在 1970~2100 年、纬度绝对值不超过 90 度的域内，高度角误差优于 0.5 度。
 *   本件不做大气折射修正（折射在地平线附近可达 0.5 度），日出日落判据请以
 *   bSunUp 为「几何高度角为正」而非「可见日面出地平」。
 * 修订历史 (Revision)   :
 *   2026-11-15  v1.0.0  首版入库（R12 · Level 0 DL_MathData 天文钟族）
 *============================================================================*)
FUNCTION FC_DL_SolarPositionCalc : REAL
VAR_INPUT
    nYear        : INT;                  // 年 [年]，域 1970~2100 / Year, 1970..2100
    nMonth       : INT;                  // 月 [月]，域 1~12 / Month, 1..12
    nDay         : INT;                  // 日 [日]，域 1~31，按当月实际天数校验 / Day, 1..31, checked against the month
    nHour        : INT;                  // 时 [h]，域 0~23，本地标准时 / Hour, local standard time
    nMinute      : INT;                  // 分 [min]，域 0~59 / Minute, 0..59
    fLatitude    : REAL;                 // 纬度 [度]，北纬为正，域 −90~90 / Latitude in degrees, north positive
    fLongitude   : REAL;                 // 经度 [度]，东经为正，域 −180~180 / Longitude in degrees, east positive
    nUtcOffsetMin : INT := 480;          // 本地时区偏移 [min]，东八区 = 480 / Time zone offset in minutes
END_VAR
VAR_OUTPUT
    fDeclination : REAL;                 // 太阳赤纬 [度]，约 −23.45~+23.45 / Solar declination in degrees
    fHourAngle   : REAL;                 // 时角 [度]，正午为 0，下午为正 / Hour angle in degrees
    fElevation   : REAL;                 // 太阳高度角 [度]，地平线上为正 / Solar elevation in degrees
    fAzimuth     : REAL;                 // 方位角 [度]，正北 0 顺时针增 / Azimuth clockwise from north
    fEquationOfTime : REAL;              // 均时差 [min] / Equation of time in minutes
    bSunUp       : BOOL;                 // 高度角大于 0 = TRUE / Sun above the horizon
    uErrorId     : UDINT;                // 事件码，0 = 无事件 / Event code, zero means none
    bValid       : BOOL;                 // 日期、时区、经纬度均合法 = TRUE / All inputs legal
END_VAR
VAR
    nDoy         : INT;                  // 年内日序，1 月 1 日 = 1 [日] / Day of year, January the first is one
    fGamma       : REAL;                 // 小数年角 [rad] / Fractional year angle in radians
    fDeclRad     : REAL;                 // 赤纬中间量 [rad] / Declination in radians
    fEotMin      : REAL;                 // 均时差中间量 [min] / Equation of time intermediate
    fTstMin      : REAL;                 // 真太阳时 [min] / True solar time in minutes
    fHaDeg       : REAL;                 // 时角中间量 [度] / Hour angle intermediate in degrees
    fLatRad      : REAL;                 // 纬度 [rad] / Latitude in radians
    fSinElev     : REAL;                 // 高度角正弦中间量 [-] / Sine of the elevation
    fCosElev     : REAL;                 // 高度角余弦中间量 [-] / Cosine of the elevation
    fY           : REAL;                 // 方位角反正切分子 [-] / Azimuth arc tangent numerator
    fX           : REAL;                 // 方位角反正切分母 [-] / Azimuth arc tangent denominator
    fAzRad       : REAL;                 // 方位角中间量 [rad] / Azimuth in radians
    nDayMax      : INT;                  // 当月天数 [日] / Days in the month
    bLeap        : BOOL;                 // 闰年标志 / Leap year flag
    i            : INT;                  // 月份累加索引 [月] / Month accumulation index
    nGuard       : DINT;                 // 循环守卫 / Loop guard
END_VAR
VAR CONSTANT
    DL_RAD2DEG   : REAL := 57.29577951;  // 弧度转度 [度] / Radians to degrees
    DL_DEG2RAD   : REAL := 0.01745329;   // 度转弧度 [rad] / Degrees to radians
    DL_PI        : REAL := 3.14159265;   // 圆周率 [-] / Pi
    DL_DAYS_YEAR : REAL := 365.0;        // 平年天数 [日] / Days in a common year
    DL_TWO_PI    : REAL := 6.28318531;   // 二倍圆周率 [rad] / Two pi
    DL_HA_LIM    : REAL := 180.0;        // 时角归一上限 [度] / Hour angle normalisation bound
    DL_AZ_FULL   : REAL := 360.0;        // 方位角整圈 [度] / Full azimuth circle in degrees
    DL_SIN_LIM   : REAL := 1.0;          // 反正弦定义域边界 [-] / Arc sine domain bound
    DL_ZENITH_DEG : REAL := 89.5;        // 天顶不可辨阈值 [度] / Zenith ambiguity threshold in degrees
    DL_COS_MIN   : REAL := 0.00873;      // 天顶不可辨的余弦阈值 [-] / Cosine threshold for the zenith case
    DL_EPS       : REAL := 1.0E-6;       // 浮点判零容差 [-] / Float zero tolerance
    DL_LAT_MAX   : REAL := 90.0;         // 纬度绝对值上限 [度] / Latitude absolute bound
    DL_LON_MAX   : REAL := 180.0;        // 经度绝对值上限 [度] / Longitude absolute bound
    DL_UTC_MAX   : INT  := 840;          // 时区偏移绝对值上限 [min] / Time zone absolute bound
    DL_YEAR_MIN  : INT  := 1970;         // 年份下限 [年] / Lower year bound
    DL_YEAR_MAX  : INT  := 2100;         // 年份上限 [年] / Upper year bound
    DL_GUARD_MAX : DINT := 16;           // 循环守卫上限 [次] / Loop guard limit
END_VAR

(*------------------------------------------------------------------------------
 * 段 1｜结果预置：全部角度出口先落 0.0，早退路径不留未初始化量
 *      Safe preset: all angle outputs fall back to 0.0 on every early exit
 *-----------------------------------------------------------------------------*)
FC_DL_SolarPositionCalc := 0.0;
fDeclination    := 0.0;
fHourAngle      := 0.0;
fElevation      := 0.0;
fAzimuth        := 0.0;
fEquationOfTime := 0.0;
bSunUp          := FALSE;
uErrorId        := 16#0000_0000;
bValid          := FALSE;
nDoy            := 0;
nDayMax         := 0;
bLeap           := FALSE;
nGuard          := 0;
i               := 1;

(*------------------------------------------------------------------------------
 * 段 2｜日期时间域闸门：年月时分越界一律早退（码 0136），不做任何夹取
 *      Date and time domain gates: out of range exits with 0136, never clamped
 *-----------------------------------------------------------------------------*)
IF (nYear < DL_YEAR_MIN) OR (nYear > DL_YEAR_MAX) THEN
    uErrorId := 16#0001_0136;
    RETURN;
END_IF
IF (nMonth < 1) OR (nMonth > 12) THEN
    uErrorId := 16#0001_0136;
    RETURN;
END_IF
IF (nHour < 0) OR (nHour > 23) THEN
    uErrorId := 16#0001_0136;
    RETURN;
END_IF
IF (nMinute < 0) OR (nMinute > 59) THEN
    uErrorId := 16#0001_0136;
    RETURN;
END_IF
IF (nUtcOffsetMin < -DL_UTC_MAX) OR (nUtcOffsetMin > DL_UTC_MAX) THEN
    uErrorId := 16#0001_0136;
    RETURN;
END_IF

(*------------------------------------------------------------------------------
 * 段 3｜地理位置域闸门：写成「正向区间取反」形式，非有限值（NaN / Inf）自然被拒
 *      Geographic gates written as inverted positive ranges so NaN is rejected too
 *      NaN 参与任何比较均为假，取反后必为真，无需额外的自比较判据
 *      NaN compares false with everything, so the inverted range catches it
 *-----------------------------------------------------------------------------*)
IF NOT ((fLatitude >= -DL_LAT_MAX) AND (fLatitude <= DL_LAT_MAX)) THEN
    uErrorId := 16#0001_0136;
    RETURN;
END_IF
IF NOT ((fLongitude >= -DL_LON_MAX) AND (fLongitude <= DL_LON_MAX)) THEN
    uErrorId := 16#0001_0136;
    RETURN;
END_IF

(*------------------------------------------------------------------------------
 * 段 4｜闰年与当月天数：4 / 100 / 400 三级判定，日越界早退（码 0137）
 *      Leap year by the 4 / 100 / 400 rule, day overflow exits with 0137
 *-----------------------------------------------------------------------------*)
bLeap := ((nYear MOD 4 = 0) AND (nYear MOD 100 <> 0)) OR (nYear MOD 400 = 0);

IF nMonth = 2 THEN
    IF bLeap THEN
        nDayMax := 29;
    ELSE
        nDayMax := 28;
    END_IF
ELSIF (nMonth = 4) OR (nMonth = 6) OR (nMonth = 9) OR (nMonth = 11) THEN
    nDayMax := 30;
ELSE
    nDayMax := 31;
END_IF

IF (nDay < 1) OR (nDay > nDayMax) THEN
    uErrorId := 16#0001_0137;
    RETURN;
END_IF

(*------------------------------------------------------------------------------
 * 段 5｜年内日序：逐月累加（不查表，规避各平台常量数组初始化差异），带守卫
 *      Day of year by month accumulation with a guard, no lookup table
 *-----------------------------------------------------------------------------*)
nDoy   := nDay;
nGuard := 0;
FOR i := 1 TO (nMonth - 1) DO
    IF nGuard >= DL_GUARD_MAX THEN
        EXIT;
    END_IF
    nGuard := nGuard + 1;
    IF i = 2 THEN
        IF bLeap THEN
            nDoy := nDoy + 29;
        ELSE
            nDoy := nDoy + 28;
        END_IF
    ELSIF (i = 4) OR (i = 6) OR (i = 9) OR (i = 11) THEN
        nDoy := nDoy + 30;
    ELSE
        nDoy := nDoy + 31;
    END_IF
END_FOR

(*------------------------------------------------------------------------------
 * 段 6｜小数年角与赤纬、均时差（NOAA 公开傅里叶级数）
 *      Fractional year angle, declination and equation of time
 *-----------------------------------------------------------------------------*)
fGamma := DL_TWO_PI / DL_DAYS_YEAR * (INT_TO_REAL(nDoy - 1) + (INT_TO_REAL(nHour) - 12.0) / 24.0);

fDeclRad := 0.006918
          - 0.399912 * COS(fGamma)
          + 0.070257 * SIN(fGamma)
          - 0.006758 * COS(2.0 * fGamma)
          + 0.000907 * SIN(2.0 * fGamma)
          - 0.002697 * COS(3.0 * fGamma)
          + 0.00148  * SIN(3.0 * fGamma);
fDeclination := fDeclRad * DL_RAD2DEG;

fEotMin := 229.18 * (0.000075
        + 0.001868 * COS(fGamma)
        - 0.032077 * SIN(fGamma)
        - 0.014615 * COS(2.0 * fGamma)
        - 0.040849 * SIN(2.0 * fGamma));
fEquationOfTime := fEotMin;

(*------------------------------------------------------------------------------
 * 段 7｜真太阳时与时角：经度按每度四分钟折算，时区偏移直接扣减
 *      True solar time and hour angle: four minutes per degree of longitude
 *-----------------------------------------------------------------------------*)
fTstMin := INT_TO_REAL(nHour * 60 + nMinute) + fEotMin + 4.0 * fLongitude - INT_TO_REAL(nUtcOffsetMin);
fHaDeg  := 15.0 * (fTstMin / 60.0 - 12.0);

(* 时角归一：条件加减，禁用取模（负数取余在各平台口径不一致）*)
(* Hour angle normalisation by conditional add and subtract, never by MOD *)
nGuard := 0;
WHILE (fHaDeg > DL_HA_LIM) AND (nGuard < DL_GUARD_MAX) DO
    fHaDeg := fHaDeg - DL_AZ_FULL;
    nGuard := nGuard + 1;
END_WHILE;
WHILE (fHaDeg < -DL_HA_LIM) AND (nGuard < DL_GUARD_MAX) DO
    fHaDeg := fHaDeg + DL_AZ_FULL;
    nGuard := nGuard + 1;
END_WHILE;
fHourAngle := fHaDeg;

(*------------------------------------------------------------------------------
 * 段 8｜高度角：先钳正弦到定义域，再取反正弦，杜绝 NaN 传播
 *      Elevation: clamp the sine into the arc sine domain before calling ASIN
 *-----------------------------------------------------------------------------*)
fLatRad := fLatitude * DL_DEG2RAD;
fSinElev := SIN(fLatRad) * SIN(fDeclRad)
          + COS(fLatRad) * COS(fDeclRad) * COS(fHaDeg * DL_DEG2RAD);
fSinElev := LIMIT(-DL_SIN_LIM, fSinElev, DL_SIN_LIM);

fElevation := ASIN(fSinElev) * DL_RAD2DEG;
fCosElev   := COS(fElevation * DL_DEG2RAD);

(*------------------------------------------------------------------------------
 * 段 9｜方位角：反正切求「相对正南」的偏角，再加 180 度换算到正北起算
 *      Azimuth: arc tangent gives the offset from south, plus 180 degrees
 *      公式成立前提为赤纬绝对值不超过 23.45 度，切不可把本式复用到高赤纬天体
 *      The formula assumes a declination within 23.45 degrees, never reuse it widely
 *-----------------------------------------------------------------------------*)
fY := SIN(fHaDeg * DL_DEG2RAD);
fX := COS(fHaDeg * DL_DEG2RAD) * SIN(fLatRad) - TAN(fDeclRad) * COS(fLatRad);

IF (ABS(fX) < DL_EPS) AND (ABS(fY) < DL_EPS) THEN
    fAzRad := 0.0;
ELSE
    fAzRad := ATAN2(fY, fX);
END_IF

fAzimuth := fAzRad * DL_RAD2DEG + 180.0;

(* 天顶不可辨：高度角余弦趋零时方位角无物理意义，统一置正南 *)
(* Zenith ambiguity: the azimuth is meaningless near the zenith, forced to south *)
IF (fElevation > DL_ZENITH_DEG) OR (fCosElev < DL_COS_MIN) THEN
    fAzimuth := 180.0;
ELSE
    nGuard := 0;
    WHILE (fAzimuth < 0.0) AND (nGuard < DL_GUARD_MAX) DO
        fAzimuth := fAzimuth + DL_AZ_FULL;
        nGuard   := nGuard + 1;
    END_WHILE;
    WHILE (fAzimuth >= DL_AZ_FULL) AND (nGuard < DL_GUARD_MAX) DO
        fAzimuth := fAzimuth - DL_AZ_FULL;
        nGuard   := nGuard + 1;
    END_WHILE;
END_IF

(*------------------------------------------------------------------------------
 * 段 10｜日出判定与出口收口：几何高度角为正即视为在地平线之上
 *      Sun up verdict and output closure based on the geometric elevation
 *-----------------------------------------------------------------------------*)
bSunUp := fElevation > 0.0;
bValid := TRUE;

FC_DL_SolarPositionCalc := fElevation;
END_FUNCTION

(* ---- FC_DL_SolveLinear3.st ---- *)
(*
  ==================================================================
  组件名 Component  : FC_DL_SolveLinear3
  分类   Category   : DL_MathData
  复杂度 Complexity  : 中
  版本   Version    : 1.0.0
  功能   Purpose    : 三阶线性方程组 A·x = b 求解。部分主元高斯消元（行选
                      最大主元 + 行交换）+ 相对奇异判据（主元绝对值 < 相对
                      容差 × 系数矩阵最大绝对值判奇异）+ 非有限入参闸。
                      与 FC_DL_Matrix3Inverse 分工互引：本件直接解 Ax=b，
                      后者求显式逆矩阵。
  来源   Source     : t2-1-lgf-math（公开数值教材 clean-room）
  溯源   Origin     : 部分主元高斯消元为公开数值教材算法，clean-room 自研
                      实现，未复制任何厂商私有库源码。
  平台   Platform   : 纯 IEC 61131-3，CODESYS / TwinCAT / InoProShop 通用
  分工声明 Split     : 与 FC_DL_Matrix3Inverse 分工——Matrix3Inverse 输出显式
                      逆矩阵供多次多右端项复用；本件单次单右端项直接求解，
                      不输出逆矩阵，不做行列式出口。
  作者   Author     : 道莅代码库 · PLC 编程专家（R58）
  ------------------------------------------------------------------
  功能说明  : 四段式防御（R45）：预置 → 非有限 / 奇异域闸 → 域内消元回代 →
              结果非有限复检兜底。消元全程行交换受固定三阶界约束（无死循环
              风险）；除子均为已证非零的主元或主元相对容差护栏。
  修订记录  : 2026-11-21 v1.0.0 首次入库（R58 批 2 · 序号 5）
*)
FUNCTION FC_DL_SolveLinear3 : BOOL
VAR_IN_OUT
    aA : ARRAY[0..2, 0..2] OF LREAL; // 系数矩阵 A [混合]，消元不改写调用方副本 / the coefficient matrix A, the caller copy untouched
    afB : ARRAY[0..2] OF LREAL;      // 右端向量 b [混合] / the right hand vector b
END_VAR
VAR_OUTPUT
    afX    : ARRAY[0..2] OF LREAL; // 解向量 x [混合] / the solution vector x
    bSingular : BOOL;              // 奇异判定（相对判据命中）[-] / the singular verdict by the relative criterion
    bNonFinite: BOOL;              // 入参非有限判定 [-] / the non finite input verdict
END_VAR
VAR
    afW   : ARRAY[0..2, 0..2] OF LREAL; // 工作系数副本 [混合] / the working coefficient copy
    afR   : ARRAY[0..2] OF LREAL;       // 工作右端副本 [混合] / the working right hand copy
    nI    : DINT;   // 行遍历索引 [行] / the row loop index
    nJ    : DINT;   // 列遍历索引 [列] / the column loop index
    nK    : DINT;   // 消元内层索引 [行] / the elimination inner index
    nPiv  : DINT;   // 主元行索引 [行] / the pivot row index
    lrMaxA: LREAL;  // 系数矩阵最大绝对值 [混合] / the max absolute coefficient
    lrPiv : LREAL;  // 当前主元值 [混合] / the current pivot value
    lrTmp : LREAL;  // 交换与消元工作量 [混合] / the swap and elimination work value
    lrFac : LREAL;  // 消元因子 [无量纲] / the elimination factor
    lrSum : LREAL;  // 回代累加工作量 [混合] / the back substitution sum
END_VAR
VAR CONSTANT
    DL_SL3_REL_EPS : LREAL := 1.0E-12; // 相对奇异容差 [无量纲] / the relative singularity tolerance
END_VAR

// 段 1｜返回值与错误状态预置安全值（四段式第一段，R45）/ segment 1, preset the return and error states
FC_DL_SolveLinear3 := FALSE; // 受理标志预置假 / preset the accepted flag false
bSingular := FALSE; // 奇异标志预置假 / preset the singular flag false
bNonFinite := FALSE; // 非有限标志预置假 / preset the non finite flag false
afX[0] := 0.0; // 解向量预置零（分量一）/ preset the solution zero, the entry one
afX[1] := 0.0; // 解向量预置零（分量二）/ preset the solution zero, the entry two
afX[2] := 0.0; // 解向量预置零（分量三）/ preset the solution zero, the entry three

// 段 2｜非有限入参闸（自反双判据全覆盖 12 个量，R79 / R151）/ segment 2, the non finite input gate over all twelve entries
FOR nI := 0 TO 2 DO // 行遍历 / the row loop
    IF (afB[nI] <> afB[nI]) OR ((afB[nI] - afB[nI]) <> (afB[nI] - afB[nI])) THEN // 右端非有限 / a non finite right hand
        bNonFinite := TRUE; // 置非有限标志 / raise the non finite flag
    END_IF
    FOR nJ := 0 TO 2 DO // 列遍历 / the column loop
        IF (aA[nI, nJ] <> aA[nI, nJ]) OR ((aA[nI, nJ] - aA[nI, nJ]) <> (aA[nI, nJ] - aA[nI, nJ])) THEN // 系数非有限 / a non finite coefficient
            bNonFinite := TRUE; // 置非有限标志 / raise the non finite flag
        END_IF
    END_FOR
END_FOR
IF bNonFinite THEN // 非有限命中：返回预置安全解 / a non finite hit, return the preset safe solution
    RETURN; // 早退（解向量保持预置零）/ return early with the preset zero
END_IF

// 段 3｜工作副本装填 + 矩阵最大绝对值（相对奇异判据基准）/ segment 3, the working copies and the max absolute coefficient
lrMaxA := 0.0; // 基准预置零 / preset the base zero
FOR nI := 0 TO 2 DO // 行遍历 / the row loop
    afR[nI] := afB[nI]; // 装右端副本 / load the right hand copy
    FOR nJ := 0 TO 2 DO // 列遍历 / the column loop
        afW[nI, nJ] := aA[nI, nJ]; // 装系数副本 / load the coefficient copy
        IF ABS(aA[nI, nJ]) > lrMaxA THEN // 更新最大绝对值 / update the max absolute
            lrMaxA := ABS(aA[nI, nJ]); // 记录基准 / record the base
        END_IF
    END_FOR
END_FOR

// 段 4｜部分主元前向消元（行选最大主元 + 行交换，固定三阶界）/ segment 4, the partial pivot forward elimination
FOR nK := 0 TO 1 DO // 消元主列遍历（末列免消）/ the pivot column loop
    nPiv := nK; // 主元行预置当前行 / preset the pivot row
    lrPiv := ABS(afW[nK, nK]); // 当前主元绝对值 / the current pivot magnitude
    FOR nI := nK + 1 TO 2 DO // 候选行遍历 / the candidate row loop
        IF ABS(afW[nI, nK]) > lrPiv THEN // 更大候选主元 / a larger candidate pivot
            nPiv := nI; // 更新主元行 / update the pivot row
            lrPiv := ABS(afW[nI, nK]); // 更新主元值 / update the pivot value
        END_IF
    END_FOR
    IF lrPiv < (DL_SL3_REL_EPS * lrMaxA) THEN // 相对奇异判据命中 / the relative singularity hit
        bSingular := TRUE; // 置奇异标志 / raise the singular flag
        RETURN; // 早退（解向量保持预置零）/ return early with the preset zero
    END_IF
    IF nPiv <> nK THEN // 需要行交换 / a row swap needed
        FOR nJ := 0 TO 2 DO // 交换系数行 / swap the coefficient rows
            lrTmp := afW[nK, nJ]; // 暂存行 K / hold row K
            afW[nK, nJ] := afW[nPiv, nJ]; // 主元行上调 / the pivot row up
            afW[nPiv, nJ] := lrTmp; // 原行落位 / the old row down
        END_FOR
        lrTmp := afR[nK]; // 交换右端同行 / swap the right hand
        afR[nK] := afR[nPiv]; // 右端同步 / sync the right hand
        afR[nPiv] := lrTmp; // 右端落位 / settle the right hand
    END_IF
    FOR nI := nK + 1 TO 2 DO // 下方行消元 / eliminate the rows below
        lrFac := afW[nI, nK] / afW[nK, nK]; // 消元因子（主元已证过容差闸）/ the elimination factor
        FOR nJ := nK TO 2 DO // 行内系数更新 / update the row coefficients
            afW[nI, nJ] := afW[nI, nJ] - lrFac * afW[nK, nJ]; // 系数消元 / eliminate the coefficient
        END_FOR
        afR[nI] := afR[nI] - lrFac * afR[nK]; // 右端消元 / eliminate the right hand
    END_FOR
END_FOR
IF ABS(afW[2, 2]) < (DL_SL3_REL_EPS * lrMaxA) THEN // 末主元相对奇异复检 / the last pivot relative singularity recheck
    bSingular := TRUE; // 置奇异标志 / raise the singular flag
    RETURN; // 早退 / return early
END_IF

// 段 5｜回代求解（除子均为主元，已证过容差闸）/ segment 5, the back substitution
FOR nI := 2 TO 0 BY -1 DO // 自下而上回代（DINT 递减步进固定界）/ the upward back substitution with a fixed bound
    lrSum := afR[nI]; // 右端起算 / start from the right hand
    FOR nJ := nI + 1 TO 2 DO // 已解分量累加 / accumulate the solved entries
        lrSum := lrSum - afW[nI, nJ] * afX[nJ]; // 扣已解项 / subtract the solved term
    END_FOR
    afX[nI] := lrSum / afW[nI, nI]; // 解出本分量（主元已证）/ solve the entry
END_FOR

// 段 6｜结果非有限复检兜底（防御纵深，正常路径不可达）/ segment 6, the result recheck as defense in depth
FOR nI := 0 TO 2 DO // 分量遍历 / the entry loop
    IF (afX[nI] <> afX[nI]) OR ((afX[nI] - afX[nI]) <> (afX[nI] - afX[nI])) THEN // 解分量非有限 / a non finite solution entry
        afX[nI] := 0.0; // 分量归零兜底 / zero the entry
        FC_DL_SolveLinear3 := FALSE; // 不予受理 / refuse the acceptance
        RETURN; // 早退 / return early
    END_IF
END_FOR
FC_DL_SolveLinear3 := TRUE; // 求解受理 / accept the solution
END_FUNCTION

(* ---- FC_DL_SortIndexLReal.st ---- *)
(*
  ==================================================================
  组件名 Component  : FC_DL_SortIndexLReal
  分类   Category   : DL_MathData
  前缀   Naming     : FC_DL_ ｜ b/n/u/f/t/e/st 类型前缀制（R265）
  复杂度 Complexity  : 中
  版本   Version    : 1.0.0
  功能   Purpose    : 稳定排序仅输出索引排列，不改调用方数组（只读纪律）。
  来源   Source     : self-std（公开排序语义自研，索引间接排序实现）
  平台   Platform   : 纯 IEC 61131-3（FOR / WHILE / 比较 / 数组），三平台通用
  分工声明 Split     : 与 FC_DL_PercentileLReal（百分位属主）分工——后者只读
                      求分位；本件出索引排列供上层复用，两件共用只读纪律
                      （R216 双向互引）。
  作者   Author     : 道莅代码库 · PLC 编程专家（R61）
  归属 Ownership     : 本件无 TYPE 声明；引用件类型全部 IEC 标准原生。
  ------------------------------------------------------------------
  边界 Boundary     :
                      一 稳定性判据写死下标序：比较用严格小于，相等元素保持
                         原下标先后（插入序即下标序），不交换等值对；
                      二 nCount = 0 / 1 退化直返恒等索引（aIdx[i] = i），不置码；
                      三 非有限元素判故障拒绝（NaN 与任何比较均假会静默破坏
                         排序，必须逐个点名，R272）；
                      四 索引写出前已证在 [0, nUse-1] 内，回钳量不再复判越界
                         （R241）；扫描禁裸 WHILE 死循环（计数器上界护栏）；
                      五 只读入参数组，不改调用方数据；
                      六 无状态纯函数：局部量段 1 显式预置（R254）。
  错误码   Codes    :
    16#0001_0637【信息级】计数越域已钳位（<0 早退，>256 钳位续扫）
    16#0001_0638【故障级】元素含非有限值，拒绝排序
  验收   Acceptance :
    算法已证（脚本）：未跑 ｜ 编译器已证（三平台）：未跑
    V1 值 3/1/2 → 索引 1/2/0；V2 值 2/2/1 → 索引 2/0/1（稳定性）
    V3 nCount=1 → 恒等索引 [0]；V4 含 NaN → 码 0638、bValid=FALSE
  修订记录 Revision  :
    2026-11-21  v1.0.0  R61 首版（批 2 · 序号 5）
  ==================================================================
*)
FUNCTION FC_DL_SortIndexLReal : BOOL
VAR_IN_OUT
    afValues : ARRAY[0..255] OF LREAL; // 待排序数值 [工程单位]，只读 / the values to sort, read only
END_VAR
VAR_INPUT
    nCount : DINT; // 参与排序个数 [个]，合法域 0..256 / the count, legal from zero to two hundred fifty six
END_VAR
VAR_OUTPUT
    aIdx   : ARRAY[0..255] OF DINT; // 排序后索引排列（aIdx[0] 为最小值原下标）/ the sorted index permutation
    bValid : BOOL;                  // 结果可用标志 [-] / the result usable flag
    eErr   : UDINT;                 // 错误码，0 = 正常 / the error code, zero is ok
    bError : BOOL;                  // 错误标志，故障级码置位（R45 配对）/ the error flag
END_VAR
VAR
    k      : DINT;  // 外层插入索引 [下标] / the outer insertion index
    m      : DINT;  // 内层前移索引 [下标] / the inner shifting index
    nUse   : DINT;  // 钳位后的个数 [个] / the clamped count
    nKey   : DINT;  // 待插元素原下标暂存 [下标] / the key original index in staging
    fKey   : LREAL; // 待插元素值暂存 [工程单位] / the key value in staging
    nGuard : DINT;  // 死循环护栏计数 [次] / the dead loop guard counter
END_VAR
VAR CONSTANT
    DL_SIL_NMAX : DINT := 256; // 排序容量上界 [个]，与数组容量一致 / the sort capacity aligned with the array
    DL_SIL_GMAX : DINT := 70000; // 护栏计数上界 [次]，大于最坏比较次数 / the guard bound above the worst case
END_VAR

// 段 1｜返回值与错误状态预置安全值 + 局部量显式预置（R45 / R254）/ segment 1, the preset
FC_DL_SortIndexLReal := FALSE; // 返回值预置假 / preset the return false
bValid := FALSE; // 有效标志预置假 / preset the validity false
eErr := 16#0000_0000; // 错误码预置正常 / preset the code to ok
bError := FALSE; // 错误标志预置假 / preset the error flag false
nUse := 0; // 个数预置零 / preset the count zero
nKey := 0; // 键下标预置零 / preset the key index zero
fKey := 0.0; // 键值预置零 / preset the key value zero
nGuard := 0; // 护栏预置零 / preset the guard zero
FOR k := 0 TO 255 DO // 索引数组全量预置恒等 / preset the index array to the identity
    aIdx[k] := k; // 恒等索引 / the identity index
END_FOR

// 段 2｜计数域闸（<0 早退，>256 钳位，边界二四）/ segment 2, the count gate
IF nCount < 0 THEN // 负数非法 / a negative count
    eErr := 16#0001_0637; // 信息级：计数越域已钳位 / informational, the count clamped
    bValid := TRUE; // 空排列合法（aIdx 已全量恒等）/ the empty permutation is legal
    FC_DL_SortIndexLReal := TRUE; // 返回成功 / return success
    RETURN; // 早退 / early return
END_IF
nUse := nCount; // 域内接管 / take the count
IF nUse > DL_SIL_NMAX THEN // 超容量 / above the capacity
    nUse := DL_SIL_NMAX; // 钳到容量 / clamp to the capacity
    eErr := 16#0001_0637; // 信息级：计数越域已钳位 / informational, the count clamped
END_IF

// 段 3｜非有限元素逐个点名（R272，边界三）/ segment 3, the element wise finiteness gate
FOR k := 0 TO nUse - 1 DO // 有界遍历 / the bounded traversal
    IF (afValues[k] <> afValues[k]) OR ((afValues[k] - afValues[k]) <> (afValues[k] - afValues[k])) THEN // 元素非有限 / the element is not finite
        eErr := 16#0001_0638; // 故障级：元素含非有限值 / fault grade, a non finite element
        bError := TRUE; // 置错误标志（R45 配对）/ raise the error flag
        bValid := FALSE; // 结果不可用 / the result void
        RETURN; // 早退（aIdx 保持恒等，不外泄坏排列）/ early return with the identity kept
    END_IF
END_FOR

// 段 4｜插入排序（索引间接，严格比较保稳定，边界一；护栏防死循环，边界四）/ segment 4, the stable insertion sort on the indices
FOR k := 1 TO nUse - 1 DO // 有界外层 / the bounded outer loop
    nKey := aIdx[k]; // 待插元素原下标 / the key original index
    fKey := afValues[nKey]; // 待插元素值 / the key value
    m := k - 1; // 内层从前一位置起 / the inner scan starts here
    nGuard := 0; // 护栏清零 / reset the guard
    WHILE (m >= 0) AND (afValues[aIdx[m]] > fKey) DO // 前驱更大才前移（严格大于，等值不交换，稳定性自证）/ shift while the predecessor is strictly greater
        aIdx[m + 1] := aIdx[m]; // 索引后移一位 / shift the index right
        m := m - 1; // 内层前移 / step the inner scan left
        nGuard := nGuard + 1; // 护栏计数推进 / advance the guard
        IF nGuard > DL_SIL_GMAX THEN // 护栏命中（结构性不可达兜底）/ the guard tripped, kept as a structural guard
            eErr := 16#0001_0638; // 故障级：排序失控复用非有限码前先判——此处不置码、强制收尾 / the forced stop without a new code
            m := -1; // 强制退出内层 / force the inner loop out
        END_IF
    END_WHILE
    aIdx[m + 1] := nKey; // 键落位（m+1 已证在 [0, k] 内，边界四）/ the key lands with a proven bound
END_FOR

// 段 5｜出口（nUse = 0/1 时 aIdx 已为恒等，边界二）/ segment 5, the outlet with the degenerate identity
bValid := TRUE; // 结果可用 / the result is usable
FC_DL_SortIndexLReal := TRUE; // 返回成功 / return success
END_FUNCTION

(* ---- FC_DL_SoundSpeedAirCalc.st ---- *)
//==============================================================================
// 函数：FC_DL_SoundSpeedAirCalc ｜ 中文名称：空气声速（温度/湿度函数）计算
// 所属子库：DL_MathData ｜ 版本：v1.0.0 ｜ 日期：2026-11-23
// 兼容：CODESYS V3.5+ / TwinCAT 3 / 汇川 InoProShop / Machine Expert（仅标准库
//       + 库内 FC_DL_VaporPressureSat）
// 功能描述：湿空气声速理想气体混合口径：干空气基准
//           c_dry = SQRT(1.4·287.05287·T_K)，湿度修正用混合摩尔质量法：
//           水汽摩尔分数 x_w = RH/100·p_ws(T)/p（饱和压取自族属主
//           FC_DL_VaporPressureSat，零内联 Magnus 常数），混合摩尔质量
//           M_mix = M_dry − x_w·(M_dry − M_w)，c = SQRT(γ·R_u·T_K/M_mix)。
//           简化声明：γ 固定取干空气值 1.4（湿空气 γ 略低，本简化使结果
//           偏保守偏低，超声流量/料位计前置换算用途可接受）。
// 开源溯源 (Origin)：原创实现（t1-2-oscat-building 建筑环境语义深化，公开
//           物理公式，零外部源码行，clean-room 独立编写）
// 公开接口清单：输入 fTempC / fRhPct / fPressPa；输出 fSoundSpeed / bValid
// 错误码表：纯函数无状态机码轨；无效输入经 bValid = FALSE 表达（哨兵返回
//           0.0），本件不占用 16#0001 段码位（邻件免让位）
// 状态机：N/A（纯函数，无状态，可重入）
// 边界行为：① 温度域 [-40, 60] °C、湿度域 [0, 100] %、总压域 [50000, 110000]
//           Pa，域外拒绝不外推；② 非有限输入 → 哨兵 0.0 返回；
//           ③ 委托属主件失败（含 bValid 回执，R72 口径）→ 哨兵 0.0 返回；
//           ④ M_mix 分母恒正（物理保证）仍做容差闸（防纪律豁免）。
// 修订历史：v1.0.0 2026-11-23 首版（R73 派单 · 批 2 · 序 9）
//==============================================================================

(*------------------------------------------------------------------------------
 * 调用示例：fC := FC_DL_SoundSpeedAirCalc(fTempC := 25.0, fRhPct := 60.0,
 *                                         fPressPa := 101325.0,
 *                                         fSoundSpeed => fV, bValid => bOk);
 * 注意：仅当 bValid = TRUE 时结果可进入超声仪表换算判据。
 *-----------------------------------------------------------------------------*)
FUNCTION FC_DL_SoundSpeedAirCalc : BOOL
VAR_INPUT
    fTempC    : LREAL;                 // 干球温度 [摄氏度]，域 -40..60 / Dry-bulb temperature [degC]
    fRhPct    : LREAL;                 // 相对湿度 [百分数]，域 0..100 / Relative humidity [percent]
    fPressPa  : LREAL;                 // 大气总压 [帕]，域 50000..110000 / Total pressure [Pa]
END_VAR
VAR_OUTPUT
    fSoundSpeed : LREAL;               // 空气声速 [米每秒] / Sound speed in air [m per s]
    bValid      : BOOL;                // 输出可用标志 / Outputs usable flag
    bClamped    : BOOL;                // 湿度输入越域已钳位声明（信息级，不置故障）/ RH clamped declaration, info level
END_VAR
VAR
    fTk       : LREAL;                 // 绝对温度 [开尔文] / Absolute temperature [K]
    fPwsPa    : LREAL;                 // 饱和水汽压 [帕]，属主件取得 / Saturation vapor pressure [Pa], from the owner FC
    bPwsValid : BOOL;                  // 属主件输出可用回执（R72 口径）/ Owner outputs-usable receipt, R72 style
    _bPwsClamped : BOOL;    // 属主件钳位回执（本件不消费，仅契约全回执） / Owner clamp receipt (unused, full-receipt contract)
    _nPwsErr     : UDINT;   // 属主件错误码回执 / Owner error-code receipt
    _bPwsError   : BOOL;    // 属主件故障级回执 / Owner fault-flag receipt
    fXw       : LREAL;                 // 水汽摩尔分数 [1] / Vapor mole fraction [1]
    fMixM     : LREAL;                 // 混合摩尔质量 [克每摩尔] / Mixture molar mass [g per mol]
END_VAR
VAR CONSTANT
    DL_SS_TMIN  : LREAL := -40.0;      // 温度有效下限 [摄氏度] / Temperature valid floor [degC]
    DL_SS_TMAX  : LREAL := 60.0;       // 温度有效上限 [摄氏度] / Temperature valid ceiling [degC]
    DL_SS_RHMAX : LREAL := 100.0;      // 湿度钳位上限 [百分数] / RH clamp ceiling [percent]
    DL_SS_PMIN  : LREAL := 50000.0;    // 总压有效下限 [帕] / Pressure valid floor [Pa]
    DL_SS_PMAX  : LREAL := 110000.0;   // 总压有效上限 [帕] / Pressure valid ceiling [Pa]
    DL_SS_GAMMA : LREAL := 1.4;        // 干空气比热比 [1]（简化口径声明）/ Dry-air heat ratio [1], simplified per header
    DL_SS_RU    : LREAL := 8.31446;    // 通用气体常数 [焦每摩尔每开尔文] / Universal gas constant [J per mol per K]
    DL_SS_MDRY  : LREAL := 28.9654;    // 干空气摩尔质量 [克每摩尔] / Dry-air molar mass [g per mol]
    DL_SS_MW    : LREAL := 18.01528;   // 水汽摩尔质量 [克每摩尔] / Water vapor molar mass [g per mol]
    DL_SS_EPS   : LREAL := 1.0E-6;     // 浮点容差与分母闸 / Float tolerance and denominator gate
    DL_SS_INF   : LREAL := 1.7976931348623157E308; // LREAL 幅值上限 / LREAL magnitude ceiling
    DL_SS_ZERO  : LREAL := 0.0;        // 无效哨兵输出值 / Sentinel output for invalid
END_VAR

// ---- 段 1｜出口默认值（纯函数无实例，无定时器/沿刷新义务）----
fSoundSpeed := DL_SS_ZERO;            // 声速哨兵零 / Sound speed sentinel zero
bValid := FALSE;                      // 缺省无效 / Invalid by default
bClamped := FALSE;                    // 钳位声明默认 FALSE / Clamped flag preset FALSE

// ---- 段 2｜输入防御：非有限值（NaN 自反判 + Inf 幅值判，R79）----
IF (fTempC <> fTempC) OR (ABS(fTempC) > DL_SS_INF)
   OR (fRhPct <> fRhPct) OR (ABS(fRhPct) > DL_SS_INF)
   OR (fPressPa <> fPressPa) OR (ABS(fPressPa) > DL_SS_INF) THEN
    FC_DL_SoundSpeedAirCalc := FALSE; // 返回无效 / Return invalid
    RETURN;                           // 哨兵零已预置（结构早退）/ sentinel preset, early exit
END_IF

// ---- 段 3｜域闸：温度/总压拒绝不外推；湿度越域钳位照算（信息级声明）----
IF (fTempC < DL_SS_TMIN) OR (fTempC > DL_SS_TMAX)
   OR (fPressPa < DL_SS_PMIN) OR (fPressPa > DL_SS_PMAX) THEN
    FC_DL_SoundSpeedAirCalc := FALSE; // 域外拒绝 / Out of range, refused
    RETURN;                           // 结构早退 / early exit
END_IF
IF (fRhPct < 0.0) OR (fRhPct > DL_SS_RHMAX) THEN
    fRhPct   := MIN(MAX(fRhPct, 0.0), DL_SS_RHMAX); // 湿度双侧钳位 / Two-sided RH clamp
    bClamped := TRUE;                 // 钳位声明置位 / Clamped flag raised
END_IF

// ---- 段 4｜饱和压委托族属主（含 bValid 回执，R72 口径；零内联 Magnus）----
IF NOT FC_DL_VaporPressureSat(fTempC := fTempC, fPvSat => fPwsPa, bClamped => _bPwsClamped,
                             eErr => _nPwsErr, bError => _bPwsError, bValid => bPwsValid) OR NOT bPwsValid THEN
    FC_DL_SoundSpeedAirCalc := FALSE; // 属主拒绝即本件拒绝 / Owner rejection propagates
    RETURN;                           // 结构早退（哨兵零已预置）/ early exit, sentinel preset
END_IF

// ---- 段 5｜声速主体：摩尔分数 → 混合摩尔质量 → 理想气体声速 ----
fTk := fTempC + 273.15;               // 摄氏度转开尔文 [开尔文] / Celsius to Kelvin [K]
fXw := (fRhPct / 100.0) * fPwsPa / fPressPa; // 水汽摩尔分数 [1] / Vapor mole fraction [1]
fXw := MIN(fXw, 1.0);                 // 摩尔分数物理上界钳位（饱和压越总压防护）/ Mole fraction clamped to 1.0
fMixM := DL_SS_MDRY - fXw * (DL_SS_MDRY - DL_SS_MW); // 混合摩尔质量 [克每摩尔] / Mixture molar mass [g per mol]
IF fMixM <= DL_SS_EPS THEN
    FC_DL_SoundSpeedAirCalc := FALSE; // 分母退化拒绝（物理上恒正，仍强制闸）/ Degenerate denominator, refused
    RETURN;                           // 结构早退 / early exit
END_IF
fSoundSpeed := SQRT(DL_SS_GAMMA * DL_SS_RU * fTk * 1000.0 / fMixM); // 声速 [米每秒]，克→千克单位换算 / Sound speed [m per s], gram to kg scale
bValid := TRUE;                       // 全部防御通过：输出可用 / Outputs usable
FC_DL_SoundSpeedAirCalc := TRUE;      // 返回 TRUE = 计算有效 / Return TRUE = computation valid
END_FUNCTION

(* ---- FC_DL_SphericalDistance.st ---- *)
(*
  FC_DL_SphericalDistance  —  球面大圆距离（haversine，纯函数）/ Great-circle distance via haversine, pure function
  分类 Category : DL_MathData
  码位 Code     : 16#05_0_05
  段位说明      : 05_0 段 04 格由 FC_DL_TrendSlopeCalc 启用，本件启用相邻 05 格（一件一码）
  版本 Version  : 1.0.0
  来源 Source   : t2-1-lgf-math — Math 分类「三角方向」待挖项落地
  溯源 Origin   : clean-room 实现，haversine 公式为公开领域数学方法，未复制任何源码行
  功能 Function : 1) 两经纬度（度）→ 球面大圆距离 [km]，haversine 公式 + ASIN 半角域钳制；
                  2) 同点分支：经纬差绝对值在容差内直接返回 0 距离（信息级码），不做三角运算；
                  3) 经纬度域钳制：纬度钳到 [-90, 90]、经度钳到 [-180, 180]，越界置信息级码并照常计算；
                  4) 服务 AGV 航点里程 / 光伏阵列地理排布 / 天文钟族等地理量场景。
  边界 Boundary : ① 角度入口（度）而非弧度，与上位地图口径一致，内部换算弧度；
                  ② 非有限输入（x <> x 判 NaN、差值自反判 Inf）直接故障码返回 0 距离；
                  ③ ASIN 域钳制：sqrt(h) 先钳到 [0,1] 再取 ASIN，杜绝浮点抖动越域；
                  ④ 反余弦域钳制声明：本实现走 ASIN 半角路径，天然域 [0,1]，无 ACOS 越域风险；
                  ⑤ 纯函数无内部状态，每拍重算；地球半径取公开常用值 6371.0088 km。
  依赖 Depends  : 无 DL_ 内部依赖，纯 IEC 61131-3（SIN/COS/ASIN/SQRT 均为标准函数）
  码表 Error codes（本件格 05_0_05，子码步进 +0x100）:
    16#0005_0105 信息级：经纬度越域已钳制，计算照常完成
    16#0005_0205 故障级：输入非有限（NaN/Inf），返回 0 距离
    16#0005_0305 信息级：同点分支（经纬差在容差内），返回 0 距离

  修订历史 Revision :
    2026-11-19  v1.0.0  R39 首版（批次 1 · 序号 3）
*)

FUNCTION FC_DL_SphericalDistance : LREAL    // 返回两点大圆距离 [km]，异常路径返回 0 / Returns distance [km], 0 on error paths
VAR_INPUT
    fLat1Deg : LREAL;                   // 点 1 纬度 [deg]，域 [-90, 90]，越界钳制 / Latitude of point 1 [deg]
    fLon1Deg : LREAL;                   // 点 1 经度 [deg]，域 [-180, 180]，越界钳制 / Longitude of point 1 [deg]
    fLat2Deg : LREAL;                   // 点 2 纬度 [deg] / Latitude of point 2 [deg]
    fLon2Deg : LREAL;                   // 点 2 经度 [deg] / Longitude of point 2 [deg]
END_VAR
VAR_OUTPUT
    bClamped : BOOL;                    // 本次输入发生越域钳位 / Inputs were clamped this call
    bSamePt  : BOOL;                    // 同点分支命中 / Same-point branch hit
    uErrorId : UDINT;                   // 事件码，0 = 无事件（本件码均为单次调用瞬时，无锁存）/ Event code, transient per call
END_VAR
VAR
    fLat1    : LREAL;                   // 点 1 纬度钳制后 [deg] / Clamped latitude 1
    fLon1    : LREAL;                   // 点 1 经度钳制后 [deg] / Clamped longitude 1
    fLat2    : LREAL;                   // 点 2 纬度钳制后 [deg] / Clamped latitude 2
    fLon2    : LREAL;                   // 点 2 经度钳制后 [deg] / Clamped longitude 2
    fPhi1    : LREAL;                   // 点 1 纬度弧度 [rad] / Latitude 1 in radians
    fPhi2    : LREAL;                   // 点 2 纬度弧度 [rad] / Latitude 2 in radians
    fDPhi    : LREAL;                   // 纬差弧度 [rad] / Latitude delta in radians
    fDLam    : LREAL;                   // 经差弧度 [rad] / Longitude delta in radians
    fSinDPhi : LREAL;                   // sin(纬差/2) 工作量 / sin of half latitude delta
    fSinDLam : LREAL;                   // sin(经差/2) 工作量 / sin of half longitude delta
    fH       : LREAL;                   // haversine 半角量 h = a，域 [0,1] 钳制后 / Haversine half-chord term, clamped to [0,1]
    fDLat    : LREAL;                   // 纬差 [deg]（同点判据用）/ Latitude delta [deg] for the same-point test
    fDLon    : LREAL;                   // 经差 [deg]（同点判据用）/ Longitude delta [deg] for the same-point test
END_VAR
VAR CONSTANT
    DL_SPH_LAT_MAX  : LREAL := 90.0;        // 纬度域上限 [deg] / Latitude domain bound
    DL_SPH_LON_MAX  : LREAL := 180.0;       // 经度域上限 [deg] / Longitude domain bound
    DL_SPH_INF_CAP  : LREAL := 1.0E30;      // 非有限值筛查幅值上限 / Non-finite magnitude screening cap
    DL_SPH_DEG2RAD  : LREAL := 0.017453292519943295;   // 度转弧度系数 π/180 [rad/deg] / Degrees to radians factor
    DL_SPH_R_EARTH  : LREAL := 6371.0088;   // 地球平均半径 [km]，公开常用值 / Mean Earth radius [km]
    DL_SPH_SAME_EPS : LREAL := 1.0E-9;      // 同点判据容差 [deg] / Same-point tolerance [deg]
    DL_SPH_ZERO     : LREAL := 0.0;         // 零距离常量 [km] / Zero distance constant
END_VAR

(* —— 段 1｜输出安全预置：任何异常路径返回 0 距离 —— *)
(* Stage 1, safe preset: every error path returns zero *)
FC_DL_SphericalDistance := 0.0;
bClamped := FALSE;
bSamePt  := FALSE;
uErrorId := 16#0005_0205;               // 缺省非有限故障码，通过路径末尾改写 / Default non-finite code, rewritten on success

(* —— 段 2｜非有限筛查（x<>x 判 NaN、差值自反判 Inf、幅值兜底） —— *)
(* Stage 2, non-finite screening *)
IF (fLat1Deg <> fLat1Deg) OR (ABS(fLat1Deg) > DL_SPH_INF_CAP) OR ((fLat1Deg - fLat1Deg) <> 0.0)
   OR (fLon1Deg <> fLon1Deg) OR (ABS(fLon1Deg) > DL_SPH_INF_CAP) OR ((fLon1Deg - fLon1Deg) <> 0.0)
   OR (fLat2Deg <> fLat2Deg) OR (ABS(fLat2Deg) > DL_SPH_INF_CAP) OR ((fLat2Deg - fLat2Deg) <> 0.0)
   OR (fLon2Deg <> fLon2Deg) OR (ABS(fLon2Deg) > DL_SPH_INF_CAP) OR ((fLon2Deg - fLon2Deg) <> 0.0) THEN
    RETURN;                             // 非有限输入：0 距离返回（预置码 0205 已在） / Non-finite input, return zero
END_IF

(* —— 段 3｜同点分支（容差内直接零距离，不做三角运算） —— *)
(* Stage 3, same-point branch *)
fDLat := fLat2Deg - fLat1Deg;
fDLon := fLon2Deg - fLon1Deg;
IF (ABS(fDLat) < DL_SPH_SAME_EPS) AND (ABS(fDLon) < DL_SPH_SAME_EPS) THEN
    bSamePt  := TRUE;
    uErrorId := 16#0005_0305;           // 信息级：同点零距
    RETURN;                             // 返回 0 距离（预置值）/ Return zero distance
END_IF

(* —— 段 4｜经纬度域钳制（越界置信息码并照常计算） —— *)
(* Stage 4, domain clamping *)
fLat1 := MIN(DL_SPH_LAT_MAX, MAX(-DL_SPH_LAT_MAX, fLat1Deg));
fLon1 := MIN(DL_SPH_LON_MAX, MAX(-DL_SPH_LON_MAX, fLon1Deg));
fLat2 := MIN(DL_SPH_LAT_MAX, MAX(-DL_SPH_LAT_MAX, fLat2Deg));
fLon2 := MIN(DL_SPH_LON_MAX, MAX(-DL_SPH_LON_MAX, fLon2Deg));
IF (fLat1 <> fLat1Deg) OR (fLon1 <> fLon1Deg) OR (fLat2 <> fLat2Deg) OR (fLon2 <> fLon2Deg) THEN
    bClamped := TRUE;
    uErrorId := 16#0005_0105;           // 信息级：越域钳制，计算照常
END_IF

(* —— 段 5｜haversine 主体（度转弧度，半角正弦构造） —— *)
(* Stage 5, haversine core *)
fPhi1    := fLat1 * DL_SPH_DEG2RAD;
fPhi2    := fLat2 * DL_SPH_DEG2RAD;
fDPhi    := (fLat2 - fLat1) * DL_SPH_DEG2RAD;
fDLam    := (fLon2 - fLon1) * DL_SPH_DEG2RAD;
fSinDPhi := SIN(fDPhi * 0.5);
fSinDLam := SIN(fDLam * 0.5);
fH := fSinDPhi * fSinDPhi + COS(fPhi1) * COS(fPhi2) * fSinDLam * fSinDLam;   // h = sin²(Δφ/2) + cosφ1·cosφ2·sin²(Δλ/2)
IF fH < 0.0 THEN
    fH := 0.0;                          // 浮点抖动下限钳位 / Clamp numerical noise below zero
END_IF
IF fH > 1.0 THEN
    fH := 1.0;                          // ASIN 域钳制（上限）：杜绝越域 / ASIN domain clamp upper
END_IF

(* —— 段 6｜距离合成：d = 2R·asin(sqrt(h))（h 已钳 [0,1]，无越域） —— *)
(* Stage 6, distance assembly *)
FC_DL_SphericalDistance := 2.0 * DL_SPH_R_EARTH * ASIN(SQRT(fH));
uErrorId := 16#0000_0000;               // 正常路径无事件 / No event on the normal path
IF bClamped THEN
    uErrorId := 16#0005_0105;           // 钳制信息码还原（正常距离照常返回）/ Restore clamp info code
END_IF

END_FUNCTION

(* ---- FC_DL_SputterDepositionRateCalc.st ---- *)
(*
  DL Factory R88 | FC_DL_SputterDepositionRateCalc
  功能：按工程简化式算溅射沉积速率 r=Y·P/(A·ρ)（Y 为含产额与几何折算的综合系数），并按带宽判合格
  开源溯源：无（clean-room 自研，依据公开工艺公式 溅射速率 r∝溅射产额×功率/(靶面积×密度)，许可证=MIT，借鉴点=公式结构）
  规则：R1-R16 全遵守；R88 简单件标量形（纯标量入参出参，无循环体、无方法、无属性、无数组）
*)
FUNCTION FC_DL_SputterDepositionRateCalc : REAL
VAR_INPUT
    fSputterYield : REAL := 2.5; // 综合速率系数 Y（含溅射产额/几何/单位折算） [-] / lumped rate coefficient [-]
    fPowerKW : REAL := 5.0; // 靶面输入功率 P [kW] / target input power [kW]
    fTargetAreaCm2 : REAL := 300.0; // 靶材有效溅射面积 A [cm²] / effective target area [cm^2]
    fDensityGcm3 : REAL := 10.2; // 靶材密度 ρ（铜 8.96，钼 10.2，铝 2.70） [g/cm³] / target density [g/cm^3]
    fMinNmMin : REAL := 10.0; // 速率允许下限（工艺带宽） [nm/min] / lower rate band [nm/min]
    fMaxNmMin : REAL := 200.0; // 速率允许上限（工艺带宽） [nm/min] / upper rate band [nm/min]
END_VAR
VAR_OUTPUT
    fRateNmMin : REAL; // 沉积速率 r [nm/min] / deposition rate [nm/min]
    xInBand : BOOL; // TRUE=速率落在允许带宽内 [-] / TRUE when inside the band [-]
END_VAR
VAR
    fDenom : REAL; // 分母 A·ρ（除零判据，单位 g/cm） [-] / denominator, the divisor [-]
    fNum : REAL; // 分子 Y·P [kW] / numerator [kW]
END_VAR

// 段 1｜出口预置
FC_DL_SputterDepositionRateCalc := -1.0; // 哨兵返回 -1（无效） [-] / sentinel return -1, invalid [-]
fRateNmMin := 0.0; // 沉积速率预置零 [nm/min] / rate preset zero [nm/min]
xInBand := FALSE; // 带宽位预置 FALSE（未判定前不认合格） [-] / band flag preset false [-]

// 段 2｜非有限拦截 + 域闸
IF NOT (fSputterYield > -1.0E30 AND fSputterYield < 1.0E30) OR NOT (fPowerKW > -1.0E30 AND fPowerKW < 1.0E30) OR NOT (fTargetAreaCm2 > -1.0E30 AND fTargetAreaCm2 < 1.0E30) THEN
    RETURN; // 综合系数/功率/靶面积任一非有限即拒算 [-] / any non finite input rejected [-]
END_IF
IF NOT (fDensityGcm3 > -1.0E30 AND fDensityGcm3 < 1.0E30) OR NOT (fMinNmMin > -1.0E30 AND fMinNmMin < 1.0E30) OR NOT (fMaxNmMin > -1.0E30 AND fMaxNmMin < 1.0E30) THEN
    RETURN; // 密度/带宽上下限任一非有限则判据静默失效，故先拦 [-] / these pins must be finite [-]
END_IF
IF fSputterYield <= 0.0 OR fPowerKW < 0.0 OR fTargetAreaCm2 < 1.0E-9 OR fDensityGcm3 < 1.0E-9 THEN
    RETURN; // 综合系数正域闸 + 功率非负闸 + 面积/密度正域闸（分母不得为零） [-] / positive gates
END_IF
IF fMinNmMin <= 0.0 OR fMaxNmMin <= fMinNmMin THEN
    RETURN; // 带宽自洽闸：下限须为正、上限须严格大于下限 [nm/min] / band consistency gate [nm/min]
END_IF

// 段 3｜计算（工程简化：不计靶面侵蚀不均、挡板遮挡与基片距离修正）
fNum := fSputterYield * fPowerKW; // [-] × kW = kW，分子合成 [kW] / [-] x [kW] = [kW]
fDenom := fTargetAreaCm2 * fDensityGcm3; // cm² × g/cm³ = g/cm，分母合成 [-] / [g/cm^3 x cm^2]
IF fDenom < 1.0E-9 THEN
    RETURN; // 除法前分母闸：A·ρ 必须大于 1E-9 才可作除数 [-] / denominator gate before the division [-]
END_IF
fRateNmMin := fNum / fDenom; // 综合系数已含单位折算，商即 nm/min [nm/min] / rate [nm/min]

// 段 4｜判定与饱和
IF NOT (fRateNmMin > -1.0E30 AND fRateNmMin < 1.0E30) THEN
    RETURN; // 结果非有限再拦一次 [-] / re-check the result for finiteness [-]
END_IF
xInBand := (fRateNmMin >= fMinNmMin) AND (fRateNmMin <= fMaxNmMin); // 双侧闭区间直比 [nm/min] / closed two sided band compare [nm/min]

// 段 5｜出口自检
IF fRateNmMin < 0.0 THEN
    RETURN; // 出口自检：速率不得为负（负值说明功率符号错） [nm/min] / rate must not be negative [nm/min]
END_IF
FC_DL_SputterDepositionRateCalc := fRateNmMin; // 返回沉积速率 [nm/min] / return the deposition rate [nm/min]
END_FUNCTION

(* ---- FC_DL_SqrtEx.st ---- *)
(*==============================================================================
 * 组件名称 (Component)  : FC_DL_SqrtEx
 * 所属子库 (Sublibrary) : DL_MathData
 * 当前版本 (Version)    : 1.0.0
 * 兼容性   (Platform)   : CODESYS 3.5 / TwinCAT 3 / 汇川 InoProShop / Machine Expert
 *                         仅依赖 Standard.library 的 SQRT 内建函数，
 *                         不重实现开方内核，无厂商数学方言依赖
 * 功能一句话 (Summary)  : 平方根防御包装：负数与非有限输入域闸门先行，
 *                         域内委托内建 SQRT，绝不向下游输出 NaN。
 * 功能描述 (Function)   : 对被开方数 fX 求平方根。定义域闸门先行写死：
 *                         fX 非有限（NaN 用 x <> x 判据、无穷用 ABS(x) 超
 *                         有限性上界判据，均为库内既有写法）或 fX < 0 时
 *                         不调内建、返回 0.0 并置码；域内（fX >= 0 且有限）
 *                         委托内建 SQRT，结果再做一次非有限复检兜底。
 * 溯源     (Origin)     : IEC 61131-3 标准语义的道莅防御性实现
 *                         （接口语义由 IEC 61131-3 定义，clean-room 重写，
 *                         参考公开标准条款）
 * 码位     (Diag Codes) : 故障级 16#0001_0227（本件独占）：
 *                           fX < 0 域外，负数开方在 IEEE 754 下产生 NaN——
 *                           本库统一为「0.0 + 故障码」策略，NaN 绝不穿透到
 *                           下游联锁（与 IEEE 默认行为的差异点，见防御声明①）；
 *                         信息级 16#0001_015A（本件独占）：
 *                           输入或输出非有限（NaN / 无穷）拦截。
 * 类型裁定 (Type Note)  : 码位段 16#0001_xxxx 为全库共享 32 位段，WORD 容量不足，
 *                         故 eErr 采用 UDINT 承载（与库内 uErrorId : UDINT 惯例
 *                         一致，沿 R14 批 3 同一裁定）。
 * 依赖     (Depends)    : 无 DL_ 内部依赖；Standard.library: SQRT / ABS
 * 红线自检 (Redline)    : R1 ✓ 零全局变量与外部变量引用 ｜ R2 ✓ 零物理 IO 地址直写
 *                         R3 ✓ 纯 IEC 61131-3 ｜ R4 ✓ 域闸门先行 + 结果非有限复检
 *                         R5 ✓ 全变量中英双语同行注释
 *                         R6 N/A（纯函数，无 CASE/ENUM 状态机，按批 4 口径标 N/A）
 *                         R7 N/A（FC 为纯函数，无实例调用，头注释显式说明）
 * 防御行为声明 (Defense): ① 负数开方返回 0.0 + 故障码 16#0001_0227，不产生
 *                           NaN——IEEE 754 下 SQRT(-x) = NaN，NaN 会沿调用链
 *                           静默污染下游滤波与比较，本库以显式码替代毒值；
 *                         ② 非有限复检先行：NaN 判据 fX <> fX（NaN 与任何值
 *                           包括自身比较均为不等，库内既有写法）、无穷判据
 *                           ABS(fX) > 1.0E308，命中即不调内建、早退返回 0.0；
 *                         ③ 域内委托内建 SQRT 内核，结果非有限复检兜底
 *                           （防御纵深，正常域内不可能触发）；
 *                         ④ fX = 0 为合法输入，SQRT(0) = 0 直通不置码；
 *                         ⑤ 1.0E308 有限性上界提为只读常量，禁魔法数；
 *                         ⑥ 浮点全程不用等号直比判数值相等，仅用 < > 与
 *                           NaN 自不等判据，符合浮点容差红线口径。
 * 修订历史 (Revision)   :
 *   2026-11-16  v1.0.0  首版入库（R14 批 4 · T0 快车道）
 *============================================================================*)
FUNCTION FC_DL_SqrtEx : LREAL
VAR_INPUT
    fX : LREAL; // 被开方数 [无量纲]，须 >= 0 且有限 / Radicand [dimensionless], must be >= 0 and finite
END_VAR
VAR_OUTPUT
    eErr : UDINT; // 错误码，16#0001_0227=负数域外，16#0001_015A=非有限拦截，0=无事件 / Error code, 16#0001_0227=negative domain, 16#0001_015A=non-finite interception, 0=no event
END_VAR
VAR CONSTANT
    DL_SQ_FINITE : LREAL := 1.0E308; // 有限性上界 [无量纲]，超界判无穷（库内既有写法）/ Finiteness bound, values beyond treated as infinity (library idiom)
END_VAR

(*------------------------------------------------------------------------------
 * 段 1｜返回值与错误码预置：先归零，任何早退路径都不会留下脏码
 *      Preset return value and error code so no early-exit path leaves a stale code
 *-----------------------------------------------------------------------------*)
FC_DL_SqrtEx := 0.0;   // 返回值预置 0.0（安全值，绝不输出 NaN）/ Preset return to 0.0 (safe value, never NaN)
eErr         := 16#0000_0000;   // 错误码预置无事件 / Preset error code to no event

(*------------------------------------------------------------------------------
 * 段 2｜非有限复检先行（防御声明②）：NaN 与无穷一律不进内建内核
 *      Non-finite recheck first (defense note 2): NaN and infinity never reach
 *      the built-in kernel
 *-----------------------------------------------------------------------------*)
IF (fX <> fX) OR (ABS(fX) > DL_SQ_FINITE) THEN
    eErr := 16#0001_015A;   // 信息码：输入非有限（NaN / 无穷），拦截早退 / Informational: non-finite input (NaN or infinity), intercepted
    RETURN;                 // 返回预置安全值 0.0 / Return preset safe value 0.0
END_IF

(*------------------------------------------------------------------------------
 * 段 3｜定义域闸门（防御声明①）：fX < 0 域外，返回 0.0 + 故障码，
 *      杜绝 IEEE 默认的 NaN 穿透（联锁回路毒值）
 *      Domain gate (defense note 1): negative input returns 0.0 with fault code,
 *      IEEE NaN propagation to downstream interlocks is eliminated
 *-----------------------------------------------------------------------------*)
IF fX < 0.0 THEN
    eErr := 16#0001_0227;   // 故障码：负数开方域外，返回安全值 0.0 / Fault: negative radicand out of domain, safe value 0.0 returned
    RETURN;                 // 返回预置安全值 0.0，不产生 NaN / Return preset safe value 0.0, no NaN produced
END_IF

(*------------------------------------------------------------------------------
 * 段 4｜域内委托内建内核（防御声明③④⑤）：fX >= 0 且有限，
 *      SQRT(0) = 0 合法直通；结果非有限复检兜底（防御纵深）
 *      In-domain delegation to the built-in kernel (defense notes 3 to 5):
 *      SQRT(0) = 0 passes legally; result recheck is defense in depth
 *-----------------------------------------------------------------------------*)
FC_DL_SqrtEx := SQRT(fX);   // 委托内建 SQRT 内核，不自实现开方 / Delegate to the built-in SQRT kernel, no re-implementation

(*------------------------------------------------------------------------------
 * 段 5｜结果非有限复检（防御声明③）：域内正常不可能触发，兜底拦截
 *      Result finiteness recheck (defense note 3): unreachable in the normal
 *      domain, kept as a bottom-line interception
 *-----------------------------------------------------------------------------*)
IF (FC_DL_SqrtEx <> FC_DL_SqrtEx) OR (ABS(FC_DL_SqrtEx) > DL_SQ_FINITE) THEN
    FC_DL_SqrtEx := 0.0;    // 兜底安全值 0.0 / Bottom-line safe value 0.0
    eErr := 16#0001_015A;   // 信息码：结果非有限拦截 / Informational: non-finite result intercepted
END_IF
END_FUNCTION

(* ---- FC_DL_StatsCoeffVarCalc.st ---- *)
(*==============================================================================
 * 组件名称 : FC_DL_StatsCoeffVarCalc ｜ 子库 : DL_MathData ｜ v1.0.1 ｜ 2026-11-24
 * 平台     : CODESYS 3.5 / TwinCAT 3 / InoProShop / Machine Expert（纯 IEC，无厂商库）
 * 功能简介 : 变异系数 CV = σ / |μ| × 100 [%]，即标准差相对均值的离散度，用于跨量纲比较
 *            工艺稳定性（灌装量、片厚、温度均匀性等）。
 * 契约     : |fMean| ≥ 1.0E-9 且 fStd ≥ 0 且入参有限 → 返回 CV [%]、bValid := TRUE；
 *            |fMean| < 1.0E-9（近零均值下 CV 无意义，商发散）→ 返回 0、bError := TRUE；
 *            fStd < 0（标准差不可能为负，属组态/上游故障，按 0 口径返回 0）→ 同上置故障；
 *            入参非有限 → 返回 0、bError := TRUE。
 * 依赖     : 无 DL_ 内部依赖（R16 自足实现），仅用标准库 ABS
 * 错误码   : R297 零码位范式：eErr 恒 0，仅以 bError / bValid 表达
 * 红线自检 : R1 零全局 R2 零%I/%Q R3 纯IEC R4 除零前置（|μ| ≥ 1.0E-9）+ 非有限拦截 + 无 = 比较
 *            R5 双语注释 R6 N/A（无状态机）R7 N/A（无定时器/沿实例）
 *            R10 无类型转换 R11 全声明行分号 R15 标识符零保留字冲突
 * 遗留假设 : 分母取 |μ| 绝对值，故负均值同样给出正的离散百分比；CV 量纲为 %（已乘 100）；
 *            近零阈值 1.0E-9 与全库统一容差口径一致；标准差为负时「按 0 处理」的出口值
 *            同样是 0，但 bError 置位以示上游异常，二者靠 bError / bValid 区分。
 * 修订历史 : 2026-11-24 R79-B 首版（统计族 1/2）
 *============================================================================*)
FUNCTION FC_DL_StatsCoeffVarCalc : LREAL
VAR_INPUT
    fMean : LREAL := 0.0; // 样本均值 μ，可负 [工程单位] / the sample mean, negative allowed
    fStd  : LREAL := 0.0; // 样本标准差 σ，须 ≥ 0 [工程单位] / the sample standard deviation, must be non negative
END_VAR
VAR_OUTPUT
    eErr   : UDINT; // 错误码，零码位范式恒 0 / error id, always zero under the zero-code rule
    bError : BOOL;  // 近零均值、负标准差或非有限入参时为真 / TRUE on a near zero mean, a negative deviation or a non finite input
    bValid : BOOL;  // 返回值可用标志 / TRUE when the return value is usable
END_VAR
VAR CONSTANT
    DL_FIN     : LREAL := 1.0E30;  // 有限性判据上界（R477 范式：ABS(x)>FIN 判 Inf，禁用 x-x 差判）/ finiteness ceiling, ABS(x)>FIN flags Inf
    DL_ZERO : LREAL := 0.0;    // 实数零哨兵 [工程单位] / the real zero sentinel
    DL_MIN  : LREAL := 1.0E-9; // 近零均值判定阈值，全库统一容差 [工程单位] / the near zero threshold shared by the library
    DL_PCT  : LREAL := 100.0;  // 百分比换算系数 [%] / the percent scaling factor
END_VAR
VAR
    fAbsMean : LREAL; // 均值绝对值，作分母 [工程单位] / the absolute mean used as the divisor
END_VAR

// 段 1｜出口预置 / segment 1, preset the exit
FC_DL_StatsCoeffVarCalc := DL_ZERO;  // 缺省零 / default zero
eErr   := 0;                         // 零码位范式 / zero-code rule
bError := FALSE;                     // 预置无故障 / preset no fault
bValid := FALSE;                     // 域闸前不认返回值 / the return value is unusable until the gates pass

// 段 2｜非有限拦截：NaN 自反判，Inf 自减判 / segment 2, the non finite gate
IF (fMean <> fMean) OR (fStd <> fStd) THEN
    bError := TRUE;                  // NaN 入参 / a NaN input
    RETURN;                          // 返回 0 / return the preset zero
END_IF
IF (ABS(fMean) > DL_FIN) OR (ABS(fStd) > DL_FIN) THEN
    bError := TRUE;                  // Inf 入参 / an infinite input
    RETURN;                          // 返回 0 / return the preset zero
END_IF

// 段 3｜负标准差域闸：σ 不可能为负，判上游故障并按 0 口径返回 / segment 3, the negative deviation gate
IF fStd < DL_ZERO THEN
    bError := TRUE;                  // 上游给错标准差 / the upstream delivered an impossible deviation
    RETURN;                          // 按 0 口径返回 0 / return zero by convention
END_IF

// 段 4｜近零均值域闸：除法前唯一必需的拦截（CV 在 μ→0 处发散）/ segment 4, the near zero mean gate
fAbsMean := ABS(fMean);              // 分母取绝对值 / the absolute mean
IF fAbsMean < DL_MIN THEN            // 禁 = 比较，用容差下界 / a tolerance bound instead of an equality test
    bError := TRUE;                  // 近零均值，CV 无意义 / the coefficient is meaningless near a zero mean
    RETURN;                          // 返回 0 / return the preset zero
END_IF

// 段 5｜出口：CV = σ / |μ| × 100 [%] / segment 5, the coefficient of variation
FC_DL_StatsCoeffVarCalc := (fStd / fAbsMean) * DL_PCT;  // 变异系数 [%] / the coefficient of variation in percent
bValid := TRUE;                      // 返回值可用 / the return value is usable
END_FUNCTION
